  movel([0.295202, -1.405507, -2.534956, -0.771926, 1.570796, 1.865998],accel_mss,speed_ms,0,blend_radius_m)
  movel([0.293033, -1.404298, -2.535858, -0.772233, 1.570796, 1.863829],accel_mss,speed_ms,0,blend_radius_m)
  movel([0.292106, -1.403830, -2.536207, -0.772352, 1.570796, 1.862902],accel_mss,speed_ms,0,blend_radius_m)
  movel([0.292065, -1.403853, -2.536190, -0.772346, 1.570796, 1.862862],accel_mss,speed_ms,0,blend_radius_m)
  movel([0.291975, -1.403947, -2.536120, -0.772322, 1.570796, 1.862771],accel_mss,speed_ms,0,blend_radius_m)
  movel([0.291907, -1.404050, -2.536043, -0.772296, 1.570796, 1.862703],accel_mss,speed_ms,0,blend_radius_m)
  movel([0.288768, -1.410063, -2.531537, -0.770789, 1.570796, 1.859564],accel_mss,speed_ms,0,blend_radius_m)
  movel([0.288784, -1.410109, -2.531502, -0.770777, 1.570796, 1.859580],accel_mss,speed_ms,0,blend_radius_m)
  movel([0.288827, -1.410120, -2.531495, -0.770775, 1.570796, 1.859623],accel_mss,speed_ms,0,blend_radius_m)
  movel([0.296146, -1.408109, -2.533007, -0.771273, 1.570796, 1.866942],accel_mss,speed_ms,0,blend_radius_m)
  movel([0.296784, -1.407940, -2.533134, -0.771315, 1.570796, 1.867580],accel_mss,speed_ms,0,blend_radius_m)
  movel([0.297418, -1.407780, -2.533254, -0.771355, 1.570796, 1.868215],accel_mss,speed_ms,0,blend_radius_m)
  movel([0.297807, -1.407689, -2.533323, -0.771378, 1.570796, 1.868604],accel_mss,speed_ms,0,blend_radius_m)
  movel([0.298196, -1.407603, -2.533387, -0.771399, 1.570796, 1.868993],accel_mss,speed_ms,0,blend_radius_m)
  movel([0.298230, -1.407602, -2.533388, -0.771399, 1.570796, 1.869026],accel_mss,speed_ms,0,blend_radius_m)
  movel([0.298257, -1.407614, -2.533378, -0.771396, 1.570796, 1.869053],accel_mss,speed_ms,0,blend_radius_m)
  movel([0.298268, -1.407641, -2.533359, -0.771390, 1.570796, 1.869065],accel_mss,speed_ms,0,blend_radius_m)
  movel([0.298265, -1.407672, -2.533335, -0.771382, 1.570796, 1.869061],accel_mss,speed_ms,0,blend_radius_m)
  movel([0.298217, -1.407806, -2.533235, -0.771348, 1.570796, 1.869013],accel_mss,speed_ms,0,blend_radius_m)
  movel([0.298155, -1.407940, -2.533134, -0.771315, 1.570796, 1.868951],accel_mss,speed_ms,0,blend_radius_m)
  movel([0.298085, -1.408074, -2.533034, -0.771281, 1.570796, 1.868881],accel_mss,speed_ms,0,blend_radius_m)
  movel([0.296508, -1.410799, -2.530982, -0.770608, 1.570796, 1.867304],accel_mss,speed_ms,0,blend_radius_m)
  movel([0.294863, -1.413645, -2.528828, -0.769916, 1.570796, 1.865659],accel_mss,speed_ms,0,blend_radius_m)
  movel([0.294838, -1.413674, -2.528806, -0.769909, 1.570796, 1.865634],accel_mss,speed_ms,0,blend_radius_m)
  movel([0.294807, -1.413696, -2.528790, -0.769904, 1.570796, 1.865603],accel_mss,speed_ms,0,blend_radius_m)
  movel([0.294773, -1.413705, -2.528783, -0.769901, 1.570796, 1.865569],accel_mss,speed_ms,0,blend_radius_m)
  movel([0.292403, -1.414377, -2.528272, -0.769740, 1.570796, 1.863199],accel_mss,speed_ms,0,blend_radius_m)
  speed_ms = 0.003
  movel([0.292403, -1.402314, -2.522404, -0.787670, 1.570796, 1.863199],accel_mss,speed_ms,0,blend_radius_m)
  speed_ms = 0.01
  movel([0.292403, -1.379125, -2.510287, -0.822977, 1.570796, 1.863199],accel_mss,speed_ms,0,blend_radius_m)
  movel([0.317529, -1.353731, -2.528171, -0.830488, 1.570796, 1.888326],accel_mss,speed_ms,0,blend_radius_m)
  movel([0.317529, -1.377341, -2.540600, -0.794448, 1.570796, 1.888326],accel_mss,speed_ms,0,blend_radius_m)
  speed_ms = 0.003
  movel([0.317529, -1.386537, -2.545131, -0.780721, 1.570796, 1.888326],accel_mss,speed_ms,0,blend_radius_m)
  speed_ms = 0.007
  movel([0.317400, -1.386449, -2.545195, -0.780745, 1.570796, 1.888196],accel_mss,speed_ms,0,blend_radius_m)
  movel([0.317282, -1.386351, -2.545265, -0.780773, 1.570796, 1.888079],accel_mss,speed_ms,0,blend_radius_m)
  movel([0.317179, -1.386239, -2.545346, -0.780804, 1.570796, 1.887975],accel_mss,speed_ms,0,blend_radius_m)
  movel([0.317088, -1.386117, -2.545434, -0.780838, 1.570796, 1.887884],accel_mss,speed_ms,0,blend_radius_m)
  movel([0.317009, -1.385985, -2.545529, -0.780875, 1.570796, 1.887805],accel_mss,speed_ms,0,blend_radius_m)
  movel([0.316947, -1.385844, -2.545630, -0.780915, 1.570796, 1.887743],accel_mss,speed_ms,0,blend_radius_m)
  movel([0.316895, -1.385687, -2.545744, -0.780959, 1.570796, 1.887691],accel_mss,speed_ms,0,blend_radius_m)
  movel([0.316856, -1.385524, -2.545861, -0.781004, 1.570796, 1.887652],accel_mss,speed_ms,0,blend_radius_m)
  movel([0.316831, -1.385353, -2.545983, -0.781052, 1.570796, 1.887627],accel_mss,speed_ms,0,blend_radius_m)
  movel([0.316820, -1.385175, -2.546111, -0.781102, 1.570796, 1.887616],accel_mss,speed_ms,0,blend_radius_m)
  movel([0.316821, -1.384994, -2.546242, -0.781153, 1.570796, 1.887617],accel_mss,speed_ms,0,blend_radius_m)
  movel([0.316837, -1.384809, -2.546374, -0.781205, 1.570796, 1.887633],accel_mss,speed_ms,0,blend_radius_m)
  movel([0.316871, -1.384610, -2.546517, -0.781261, 1.570796, 1.887668],accel_mss,speed_ms,0,blend_radius_m)
  movel([0.316923, -1.384407, -2.546663, -0.781318, 1.570796, 1.887719],accel_mss,speed_ms,0,blend_radius_m)
  movel([0.316994, -1.384201, -2.546811, -0.781377, 1.570796, 1.887790],accel_mss,speed_ms,0,blend_radius_m)
  movel([0.317085, -1.383995, -2.546959, -0.781435, 1.570796, 1.887881],accel_mss,speed_ms,0,blend_radius_m)
  movel([0.317196, -1.383778, -2.547115, -0.781496, 1.570796, 1.887992],accel_mss,speed_ms,0,blend_radius_m)
  movel([0.317324, -1.383562, -2.547269, -0.781557, 1.570796, 1.888120],accel_mss,speed_ms,0,blend_radius_m)
  movel([0.317466, -1.383347, -2.547423, -0.781618, 1.570796, 1.888262],accel_mss,speed_ms,0,blend_radius_m)
  movel([0.317621, -1.383138, -2.547573, -0.781678, 1.570796, 1.888418],accel_mss,speed_ms,0,blend_radius_m)
  movel([0.317789, -1.382934, -2.547719, -0.781736, 1.570796, 1.888585],accel_mss,speed_ms,0,blend_radius_m)
  movel([0.317971, -1.382735, -2.547862, -0.781792, 1.570796, 1.888767],accel_mss,speed_ms,0,blend_radius_m)
  movel([0.318163, -1.382544, -2.547998, -0.781847, 1.570796, 1.888959],accel_mss,speed_ms,0,blend_radius_m)
  movel([0.318364, -1.382361, -2.548129, -0.781899, 1.570796, 1.889161],accel_mss,speed_ms,0,blend_radius_m)
  movel([0.318563, -1.382197, -2.548246, -0.781946, 1.570796, 1.889360],accel_mss,speed_ms,0,blend_radius_m)
  movel([0.318773, -1.382043, -2.548356, -0.781989, 1.570796, 1.889569],accel_mss,speed_ms,0,blend_radius_m)
  movel([0.318988, -1.381904, -2.548455, -0.782029, 1.570796, 1.889784],accel_mss,speed_ms,0,blend_radius_m)
  movel([0.319211, -1.381778, -2.548546, -0.782065, 1.570796, 1.890007],accel_mss,speed_ms,0,blend_radius_m)
  movel([0.319370, -1.381698, -2.548603, -0.782088, 1.570796, 1.890166],accel_mss,speed_ms,0,blend_radius_m)
  movel([0.319528, -1.381626, -2.548654, -0.782109, 1.570796, 1.890324],accel_mss,speed_ms,0,blend_radius_m)
  movel([0.319666, -1.381574, -2.548691, -0.782124, 1.570796, 1.890463],accel_mss,speed_ms,0,blend_radius_m)
  movel([0.319802, -1.381535, -2.548719, -0.782135, 1.570796, 1.890598],accel_mss,speed_ms,0,blend_radius_m)
  movel([0.319954, -1.381503, -2.548742, -0.782144, 1.570796, 1.890750],accel_mss,speed_ms,0,blend_radius_m)
  movel([0.320103, -1.381485, -2.548755, -0.782149, 1.570796, 1.890899],accel_mss,speed_ms,0,blend_radius_m)
  movel([0.320317, -1.381467, -2.548768, -0.782154, 1.570796, 1.891114],accel_mss,speed_ms,0,blend_radius_m)
  movel([0.320529, -1.381457, -2.548775, -0.782157, 1.570796, 1.891326],accel_mss,speed_ms,0,blend_radius_m)
  movel([0.320739, -1.381453, -2.548778, -0.782158, 1.570796, 1.891535],accel_mss,speed_ms,0,blend_radius_m)
  movel([0.320944, -1.381456, -2.548776, -0.782157, 1.570796, 1.891740],accel_mss,speed_ms,0,blend_radius_m)
  movel([0.321088, -1.381466, -2.548768, -0.782154, 1.570796, 1.891884],accel_mss,speed_ms,0,blend_radius_m)
  movel([0.321225, -1.381490, -2.548751, -0.782148, 1.570796, 1.892021],accel_mss,speed_ms,0,blend_radius_m)
  movel([0.321339, -1.381527, -2.548725, -0.782137, 1.570796, 1.892135],accel_mss,speed_ms,0,blend_radius_m)
  movel([0.321447, -1.381575, -2.548691, -0.782123, 1.570796, 1.892243],accel_mss,speed_ms,0,blend_radius_m)
  movel([0.321565, -1.381645, -2.548640, -0.782103, 1.570796, 1.892361],accel_mss,speed_ms,0,blend_radius_m)
  movel([0.321678, -1.381723, -2.548585, -0.782081, 1.570796, 1.892474],accel_mss,speed_ms,0,blend_radius_m)
  movel([0.321782, -1.381815, -2.548519, -0.782055, 1.570796, 1.892578],accel_mss,speed_ms,0,blend_radius_m)
  movel([0.321874, -1.381914, -2.548449, -0.782026, 1.570796, 1.892671],accel_mss,speed_ms,0,blend_radius_m)
  movel([0.321956, -1.382025, -2.548370, -0.781995, 1.570796, 1.892752],accel_mss,speed_ms,0,blend_radius_m)
  movel([0.322026, -1.382143, -2.548285, -0.781961, 1.570796, 1.892822],accel_mss,speed_ms,0,blend_radius_m)
  movel([0.322084, -1.382268, -2.548195, -0.781925, 1.570796, 1.892880],accel_mss,speed_ms,0,blend_radius_m)
  movel([0.322142, -1.382446, -2.548068, -0.781875, 1.570796, 1.892938],accel_mss,speed_ms,0,blend_radius_m)
  movel([0.322181, -1.382631, -2.547936, -0.781822, 1.570796, 1.892978],accel_mss,speed_ms,0,blend_radius_m)
  movel([0.322201, -1.382827, -2.547796, -0.781766, 1.570796, 1.892998],accel_mss,speed_ms,0,blend_radius_m)
  movel([0.322206, -1.383028, -2.547652, -0.781709, 1.570796, 1.893002],accel_mss,speed_ms,0,blend_radius_m)
  movel([0.322190, -1.383244, -2.547497, -0.781648, 1.570796, 1.892986],accel_mss,speed_ms,0,blend_radius_m)
  movel([0.322153, -1.383466, -2.547339, -0.781585, 1.570796, 1.892949],accel_mss,speed_ms,0,blend_radius_m)
  movel([0.322100, -1.383688, -2.547179, -0.781522, 1.570796, 1.892897],accel_mss,speed_ms,0,blend_radius_m)
  movel([0.322031, -1.383914, -2.547017, -0.781458, 1.570796, 1.892827],accel_mss,speed_ms,0,blend_radius_m)
  movel([0.321941, -1.384144, -2.546852, -0.781393, 1.570796, 1.892738],accel_mss,speed_ms,0,blend_radius_m)
  movel([0.321837, -1.384373, -2.546688, -0.781328, 1.570796, 1.892633],accel_mss,speed_ms,0,blend_radius_m)
  movel([0.321714, -1.384603, -2.546523, -0.781263, 1.570796, 1.892510],accel_mss,speed_ms,0,blend_radius_m)
  movel([0.321577, -1.384828, -2.546361, -0.781200, 1.570796, 1.892373],accel_mss,speed_ms,0,blend_radius_m)
  movel([0.321470, -1.384985, -2.546248, -0.781156, 1.570796, 1.892267],accel_mss,speed_ms,0,blend_radius_m)
  movel([0.321350, -1.385137, -2.546139, -0.781113, 1.570796, 1.892146],accel_mss,speed_ms,0,blend_radius_m)
  movel([0.321218, -1.385283, -2.546034, -0.781072, 1.570796, 1.892014],accel_mss,speed_ms,0,blend_radius_m)
  movel([0.321054, -1.385449, -2.545914, -0.781025, 1.570796, 1.891850],accel_mss,speed_ms,0,blend_radius_m)
  movel([0.320882, -1.385612, -2.545798, -0.780980, 1.570796, 1.891679],accel_mss,speed_ms,0,blend_radius_m)
  movel([0.320704, -1.385768, -2.545685, -0.780936, 1.570796, 1.891500],accel_mss,speed_ms,0,blend_radius_m)
  movel([0.320519, -1.385918, -2.545577, -0.780894, 1.570796, 1.891315],accel_mss,speed_ms,0,blend_radius_m)
  movel([0.320332, -1.386060, -2.545475, -0.780854, 1.570796, 1.891128],accel_mss,speed_ms,0,blend_radius_m)
  movel([0.320137, -1.386198, -2.545375, -0.780815, 1.570796, 1.890934],accel_mss,speed_ms,0,blend_radius_m)
  movel([0.319967, -1.386307, -2.545297, -0.780785, 1.570796, 1.890763],accel_mss,speed_ms,0,blend_radius_m)
  movel([0.319794, -1.386402, -2.545228, -0.780759, 1.570796, 1.890590],accel_mss,speed_ms,0,blend_radius_m)
  movel([0.319615, -1.386489, -2.545165, -0.780734, 1.570796, 1.890411],accel_mss,speed_ms,0,blend_radius_m)
  movel([0.319423, -1.386569, -2.545108, -0.780712, 1.570796, 1.890219],accel_mss,speed_ms,0,blend_radius_m)
  movel([0.319229, -1.386634, -2.545061, -0.780694, 1.570796, 1.890026],accel_mss,speed_ms,0,blend_radius_m)
  movel([0.319037, -1.386688, -2.545022, -0.780679, 1.570796, 1.889833],accel_mss,speed_ms,0,blend_radius_m)
  movel([0.318848, -1.386727, -2.544994, -0.780668, 1.570796, 1.889644],accel_mss,speed_ms,0,blend_radius_m)
  movel([0.318659, -1.386753, -2.544976, -0.780661, 1.570796, 1.889455],accel_mss,speed_ms,0,blend_radius_m)
  movel([0.318477, -1.386763, -2.544968, -0.780658, 1.570796, 1.889273],accel_mss,speed_ms,0,blend_radius_m)
  movel([0.318298, -1.386760, -2.544970, -0.780659, 1.570796, 1.889094],accel_mss,speed_ms,0,blend_radius_m)
  movel([0.318128, -1.386741, -2.544984, -0.780664, 1.570796, 1.888925],accel_mss,speed_ms,0,blend_radius_m)
  movel([0.317963, -1.386711, -2.545005, -0.780672, 1.570796, 1.888759],accel_mss,speed_ms,0,blend_radius_m)
  movel([0.317810, -1.386666, -2.545038, -0.780685, 1.570796, 1.888606],accel_mss,speed_ms,0,blend_radius_m)
  movel([0.317665, -1.386608, -2.545080, -0.780701, 1.570796, 1.888461],accel_mss,speed_ms,0,blend_radius_m)
  movel([0.317529, -1.386537, -2.545131, -0.780721, 1.570796, 1.888326],accel_mss,speed_ms,0,blend_radius_m)
  speed_ms = 0.003
  movel([0.317529, -1.389645, -2.546625, -0.776120, 1.570796, 1.888326],accel_mss,speed_ms,0,blend_radius_m)
  speed_ms = 0.007
  movel([0.317400, -1.389556, -2.546689, -0.776144, 1.570796, 1.888196],accel_mss,speed_ms,0,blend_radius_m)
  movel([0.317282, -1.389458, -2.546760, -0.776171, 1.570796, 1.888079],accel_mss,speed_ms,0,blend_radius_m)
  movel([0.317179, -1.389346, -2.546841, -0.776202, 1.570796, 1.887975],accel_mss,speed_ms,0,blend_radius_m)
  movel([0.317088, -1.389225, -2.546929, -0.776235, 1.570796, 1.887884],accel_mss,speed_ms,0,blend_radius_m)
  movel([0.317009, -1.389094, -2.547024, -0.776272, 1.570796, 1.887805],accel_mss,speed_ms,0,blend_radius_m)
  movel([0.316947, -1.388953, -2.547126, -0.776311, 1.570796, 1.887743],accel_mss,speed_ms,0,blend_radius_m)
  movel([0.316895, -1.388796, -2.547239, -0.776354, 1.570796, 1.887691],accel_mss,speed_ms,0,blend_radius_m)
  movel([0.316856, -1.388633, -2.547356, -0.776399, 1.570796, 1.887652],accel_mss,speed_ms,0,blend_radius_m)
  movel([0.316831, -1.388463, -2.547479, -0.776446, 1.570796, 1.887627],accel_mss,speed_ms,0,blend_radius_m)
  movel([0.316820, -1.388286, -2.547608, -0.776496, 1.570796, 1.887616],accel_mss,speed_ms,0,blend_radius_m)
  movel([0.316821, -1.388105, -2.547738, -0.776546, 1.570796, 1.887617],accel_mss,speed_ms,0,blend_radius_m)
  movel([0.316837, -1.387921, -2.547871, -0.776597, 1.570796, 1.887633],accel_mss,speed_ms,0,blend_radius_m)
  movel([0.316871, -1.387722, -2.548015, -0.776652, 1.570796, 1.887668],accel_mss,speed_ms,0,blend_radius_m)
  movel([0.316923, -1.387520, -2.548160, -0.776709, 1.570796, 1.887719],accel_mss,speed_ms,0,blend_radius_m)
  movel([0.316994, -1.387314, -2.548309, -0.776766, 1.570796, 1.887790],accel_mss,speed_ms,0,blend_radius_m)
  movel([0.317085, -1.387108, -2.548457, -0.776824, 1.570796, 1.887881],accel_mss,speed_ms,0,blend_radius_m)
  movel([0.317196, -1.386892, -2.548613, -0.776884, 1.570796, 1.887992],accel_mss,speed_ms,0,blend_radius_m)
  movel([0.317324, -1.386677, -2.548768, -0.776944, 1.570796, 1.888120],accel_mss,speed_ms,0,blend_radius_m)
  movel([0.317466, -1.386462, -2.548922, -0.777004, 1.570796, 1.888262],accel_mss,speed_ms,0,blend_radius_m)
  movel([0.317621, -1.386253, -2.549073, -0.777063, 1.570796, 1.888418],accel_mss,speed_ms,0,blend_radius_m)
  movel([0.317789, -1.386050, -2.549219, -0.777120, 1.570796, 1.888585],accel_mss,speed_ms,0,blend_radius_m)
  movel([0.317971, -1.385851, -2.549362, -0.777176, 1.570796, 1.888767],accel_mss,speed_ms,0,blend_radius_m)
  movel([0.318163, -1.385661, -2.549499, -0.777229, 1.570796, 1.888959],accel_mss,speed_ms,0,blend_radius_m)
  movel([0.318364, -1.385478, -2.549630, -0.777281, 1.570796, 1.889161],accel_mss,speed_ms,0,blend_radius_m)
  movel([0.318563, -1.385315, -2.549747, -0.777327, 1.570796, 1.889360],accel_mss,speed_ms,0,blend_radius_m)
  movel([0.318773, -1.385162, -2.549857, -0.777370, 1.570796, 1.889569],accel_mss,speed_ms,0,blend_radius_m)
  movel([0.318988, -1.385023, -2.549957, -0.777409, 1.570796, 1.889784],accel_mss,speed_ms,0,blend_radius_m)
  movel([0.319211, -1.384897, -2.550047, -0.777445, 1.570796, 1.890007],accel_mss,speed_ms,0,blend_radius_m)
  movel([0.319370, -1.384817, -2.550105, -0.777467, 1.570796, 1.890166],accel_mss,speed_ms,0,blend_radius_m)
  movel([0.319528, -1.384746, -2.550156, -0.777488, 1.570796, 1.890324],accel_mss,speed_ms,0,blend_radius_m)
  movel([0.319666, -1.384693, -2.550193, -0.777502, 1.570796, 1.890463],accel_mss,speed_ms,0,blend_radius_m)
  movel([0.319802, -1.384654, -2.550221, -0.777513, 1.570796, 1.890598],accel_mss,speed_ms,0,blend_radius_m)
  movel([0.319954, -1.384623, -2.550244, -0.777522, 1.570796, 1.890750],accel_mss,speed_ms,0,blend_radius_m)
  movel([0.320103, -1.384604, -2.550257, -0.777528, 1.570796, 1.890899],accel_mss,speed_ms,0,blend_radius_m)
  movel([0.320317, -1.384587, -2.550270, -0.777532, 1.570796, 1.891114],accel_mss,speed_ms,0,blend_radius_m)
  movel([0.320529, -1.384576, -2.550277, -0.777535, 1.570796, 1.891326],accel_mss,speed_ms,0,blend_radius_m)
  movel([0.320739, -1.384573, -2.550280, -0.777537, 1.570796, 1.891535],accel_mss,speed_ms,0,blend_radius_m)
  movel([0.320944, -1.384576, -2.550278, -0.777536, 1.570796, 1.891740],accel_mss,speed_ms,0,blend_radius_m)
  movel([0.321088, -1.384586, -2.550270, -0.777533, 1.570796, 1.891884],accel_mss,speed_ms,0,blend_radius_m)
  movel([0.321225, -1.384610, -2.550253, -0.777526, 1.570796, 1.892021],accel_mss,speed_ms,0,blend_radius_m)
  movel([0.321339, -1.384646, -2.550227, -0.777516, 1.570796, 1.892135],accel_mss,speed_ms,0,blend_radius_m)
  movel([0.321447, -1.384694, -2.550193, -0.777502, 1.570796, 1.892243],accel_mss,speed_ms,0,blend_radius_m)
  movel([0.321565, -1.384765, -2.550142, -0.777482, 1.570796, 1.892361],accel_mss,speed_ms,0,blend_radius_m)
  movel([0.321678, -1.384842, -2.550086, -0.777460, 1.570796, 1.892474],accel_mss,speed_ms,0,blend_radius_m)
  movel([0.321782, -1.384934, -2.550021, -0.777434, 1.570796, 1.892578],accel_mss,speed_ms,0,blend_radius_m)
  movel([0.321874, -1.385032, -2.549950, -0.777407, 1.570796, 1.892671],accel_mss,speed_ms,0,blend_radius_m)
  movel([0.321956, -1.385143, -2.549871, -0.777375, 1.570796, 1.892752],accel_mss,speed_ms,0,blend_radius_m)
  movel([0.322026, -1.385261, -2.549786, -0.777342, 1.570796, 1.892822],accel_mss,speed_ms,0,blend_radius_m)
  movel([0.322084, -1.385386, -2.549696, -0.777307, 1.570796, 1.892880],accel_mss,speed_ms,0,blend_radius_m)
  movel([0.322142, -1.385563, -2.549569, -0.777257, 1.570796, 1.892938],accel_mss,speed_ms,0,blend_radius_m)
  movel([0.322181, -1.385748, -2.549436, -0.777205, 1.570796, 1.892978],accel_mss,speed_ms,0,blend_radius_m)
  movel([0.322201, -1.385943, -2.549296, -0.777150, 1.570796, 1.892998],accel_mss,speed_ms,0,blend_radius_m)
  movel([0.322206, -1.386144, -2.549151, -0.777094, 1.570796, 1.893002],accel_mss,speed_ms,0,blend_radius_m)
  movel([0.322190, -1.386359, -2.548997, -0.777033, 1.570796, 1.892986],accel_mss,speed_ms,0,blend_radius_m)
  movel([0.322153, -1.386580, -2.548837, -0.776971, 1.570796, 1.892949],accel_mss,speed_ms,0,blend_radius_m)
  movel([0.322100, -1.386802, -2.548677, -0.776909, 1.570796, 1.892897],accel_mss,speed_ms,0,blend_radius_m)
  movel([0.322031, -1.387028, -2.548515, -0.776846, 1.570796, 1.892827],accel_mss,speed_ms,0,blend_radius_m)
  movel([0.321941, -1.387257, -2.548350, -0.776782, 1.570796, 1.892738],accel_mss,speed_ms,0,blend_radius_m)
  movel([0.321837, -1.387485, -2.548185, -0.776718, 1.570796, 1.892633],accel_mss,speed_ms,0,blend_radius_m)
  movel([0.321714, -1.387715, -2.548020, -0.776654, 1.570796, 1.892510],accel_mss,speed_ms,0,blend_radius_m)
  movel([0.321577, -1.387939, -2.547858, -0.776592, 1.570796, 1.892373],accel_mss,speed_ms,0,blend_radius_m)
  movel([0.321470, -1.388096, -2.547745, -0.776548, 1.570796, 1.892267],accel_mss,speed_ms,0,blend_radius_m)
  movel([0.321350, -1.388248, -2.547635, -0.776506, 1.570796, 1.892146],accel_mss,speed_ms,0,blend_radius_m)
  movel([0.321218, -1.388393, -2.547530, -0.776466, 1.570796, 1.892014],accel_mss,speed_ms,0,blend_radius_m)
  movel([0.321054, -1.388559, -2.547410, -0.776420, 1.570796, 1.891850],accel_mss,speed_ms,0,blend_radius_m)
  movel([0.320882, -1.388721, -2.547293, -0.776375, 1.570796, 1.891679],accel_mss,speed_ms,0,blend_radius_m)
  movel([0.320704, -1.388877, -2.547180, -0.776332, 1.570796, 1.891500],accel_mss,speed_ms,0,blend_radius_m)
  movel([0.320519, -1.389027, -2.547072, -0.776290, 1.570796, 1.891315],accel_mss,speed_ms,0,blend_radius_m)
  movel([0.320332, -1.389169, -2.546969, -0.776251, 1.570796, 1.891128],accel_mss,speed_ms,0,blend_radius_m)
  movel([0.320137, -1.389306, -2.546870, -0.776213, 1.570796, 1.890934],accel_mss,speed_ms,0,blend_radius_m)
  movel([0.319967, -1.389414, -2.546792, -0.776183, 1.570796, 1.890763],accel_mss,speed_ms,0,blend_radius_m)
  movel([0.319794, -1.389510, -2.546723, -0.776157, 1.570796, 1.890590],accel_mss,speed_ms,0,blend_radius_m)
  movel([0.319615, -1.389597, -2.546660, -0.776133, 1.570796, 1.890411],accel_mss,speed_ms,0,blend_radius_m)
  movel([0.319423, -1.389676, -2.546602, -0.776111, 1.570796, 1.890219],accel_mss,speed_ms,0,blend_radius_m)
  movel([0.319229, -1.389741, -2.546555, -0.776093, 1.570796, 1.890026],accel_mss,speed_ms,0,blend_radius_m)
  movel([0.319037, -1.389795, -2.546516, -0.776078, 1.570796, 1.889833],accel_mss,speed_ms,0,blend_radius_m)
  movel([0.318848, -1.389833, -2.546488, -0.776067, 1.570796, 1.889644],accel_mss,speed_ms,0,blend_radius_m)
  movel([0.318659, -1.389859, -2.546469, -0.776060, 1.570796, 1.889455],accel_mss,speed_ms,0,blend_radius_m)
  movel([0.318477, -1.389869, -2.546462, -0.776058, 1.570796, 1.889273],accel_mss,speed_ms,0,blend_radius_m)
  movel([0.318298, -1.389866, -2.546464, -0.776058, 1.570796, 1.889094],accel_mss,speed_ms,0,blend_radius_m)
  movel([0.318128, -1.389848, -2.546478, -0.776064, 1.570796, 1.888925],accel_mss,speed_ms,0,blend_radius_m)
  movel([0.317963, -1.389818, -2.546499, -0.776072, 1.570796, 1.888759],accel_mss,speed_ms,0,blend_radius_m)
  movel([0.317810, -1.389772, -2.546532, -0.776084, 1.570796, 1.888606],accel_mss,speed_ms,0,blend_radius_m)
  movel([0.317665, -1.389715, -2.546574, -0.776100, 1.570796, 1.888461],accel_mss,speed_ms,0,blend_radius_m)
  movel([0.317529, -1.389645, -2.546625, -0.776120, 1.570796, 1.888326],accel_mss,speed_ms,0,blend_radius_m)
  speed_ms = 0.003
  movel([0.317529, -1.377341, -2.540600, -0.794448, 1.570796, 1.888326],accel_mss,speed_ms,0,blend_radius_m)
  speed_ms = 0.01
  movel([0.317529, -1.353731, -2.528171, -0.830488, 1.570796, 1.888326],accel_mss,speed_ms,0,blend_radius_m)
  movel([0.299954, -1.366063, -2.519594, -0.826732, 1.570796, 1.870750],accel_mss,speed_ms,0,blend_radius_m)
  movel([0.299954, -1.389472, -2.531871, -0.791046, 1.570796, 1.870750],accel_mss,speed_ms,0,blend_radius_m)
  speed_ms = 0.003
  movel([0.299954, -1.398583, -2.536345, -0.777462, 1.570796, 1.870750],accel_mss,speed_ms,0,blend_radius_m)
  speed_ms = 0.007
  movel([0.299979, -1.398601, -2.536331, -0.777457, 1.570796, 1.870775],accel_mss,speed_ms,0,blend_radius_m)
  movel([0.299990, -1.398630, -2.536310, -0.777450, 1.570796, 1.870786],accel_mss,speed_ms,0,blend_radius_m)
  movel([0.299985, -1.398664, -2.536284, -0.777441, 1.570796, 1.870782],accel_mss,speed_ms,0,blend_radius_m)
  movel([0.299976, -1.398686, -2.536268, -0.777435, 1.570796, 1.870772],accel_mss,speed_ms,0,blend_radius_m)
  movel([0.299706, -1.399170, -2.535911, -0.777308, 1.570796, 1.870502],accel_mss,speed_ms,0,blend_radius_m)
  movel([0.299404, -1.399711, -2.535511, -0.777167, 1.570796, 1.870201],accel_mss,speed_ms,0,blend_radius_m)
  movel([0.299046, -1.400345, -2.535042, -0.777003, 1.570796, 1.869842],accel_mss,speed_ms,0,blend_radius_m)
  movel([0.298078, -1.402098, -2.533741, -0.776550, 1.570796, 1.868875],accel_mss,speed_ms,0,blend_radius_m)
  movel([0.298054, -1.402119, -2.533726, -0.776545, 1.570796, 1.868850],accel_mss,speed_ms,0,blend_radius_m)
  movel([0.298027, -1.402128, -2.533719, -0.776542, 1.570796, 1.868823],accel_mss,speed_ms,0,blend_radius_m)
  movel([0.298001, -1.402124, -2.533722, -0.776543, 1.570796, 1.868797],accel_mss,speed_ms,0,blend_radius_m)
  movel([0.297791, -1.402026, -2.533795, -0.776569, 1.570796, 1.868587],accel_mss,speed_ms,0,blend_radius_m)
  movel([0.297586, -1.401919, -2.533874, -0.776596, 1.570796, 1.868382],accel_mss,speed_ms,0,blend_radius_m)
  movel([0.297210, -1.401715, -2.534026, -0.776648, 1.570796, 1.868006],accel_mss,speed_ms,0,blend_radius_m)
  movel([0.296838, -1.401504, -2.534182, -0.776703, 1.570796, 1.867634],accel_mss,speed_ms,0,blend_radius_m)
  movel([0.294823, -1.400338, -2.535047, -0.777004, 1.570796, 1.865620],accel_mss,speed_ms,0,blend_radius_m)
  movel([0.291768, -1.398674, -2.536277, -0.777438, 1.570796, 1.862565],accel_mss,speed_ms,0,blend_radius_m)
  movel([0.291698, -1.398742, -2.536227, -0.777420, 1.570796, 1.862494],accel_mss,speed_ms,0,blend_radius_m)
  movel([0.291646, -1.398819, -2.536170, -0.777400, 1.570796, 1.862443],accel_mss,speed_ms,0,blend_radius_m)
  movel([0.286418, -1.408830, -2.528706, -0.774853, 1.570796, 1.857214],accel_mss,speed_ms,0,blend_radius_m)
  movel([0.286404, -1.408924, -2.528635, -0.774830, 1.570796, 1.857200],accel_mss,speed_ms,0,blend_radius_m)
  movel([0.286418, -1.408956, -2.528611, -0.774822, 1.570796, 1.857214],accel_mss,speed_ms,0,blend_radius_m)
  movel([0.286461, -1.408960, -2.528608, -0.774821, 1.570796, 1.857257],accel_mss,speed_ms,0,blend_radius_m)
  movel([0.289039, -1.408279, -2.529120, -0.774990, 1.570796, 1.859835],accel_mss,speed_ms,0,blend_radius_m)
  movel([0.292788, -1.407230, -2.529908, -0.775251, 1.570796, 1.863584],accel_mss,speed_ms,0,blend_radius_m)
  movel([0.294307, -1.406809, -2.530224, -0.775356, 1.570796, 1.865103],accel_mss,speed_ms,0,blend_radius_m)
  movel([0.295651, -1.406440, -2.530501, -0.775448, 1.570796, 1.866448],accel_mss,speed_ms,0,blend_radius_m)
  movel([0.295756, -1.406418, -2.530517, -0.775454, 1.570796, 1.866552],accel_mss,speed_ms,0,blend_radius_m)
  movel([0.295779, -1.406422, -2.530514, -0.775453, 1.570796, 1.866575],accel_mss,speed_ms,0,blend_radius_m)
  movel([0.295789, -1.406438, -2.530502, -0.775449, 1.570796, 1.866585],accel_mss,speed_ms,0,blend_radius_m)
  movel([0.295786, -1.406461, -2.530485, -0.775443, 1.570796, 1.866582],accel_mss,speed_ms,0,blend_radius_m)
  movel([0.295610, -1.406827, -2.530211, -0.775351, 1.570796, 1.866406],accel_mss,speed_ms,0,blend_radius_m)
  movel([0.295483, -1.407076, -2.530024, -0.775289, 1.570796, 1.866279],accel_mss,speed_ms,0,blend_radius_m)
  movel([0.295348, -1.407323, -2.529838, -0.775227, 1.570796, 1.866144],accel_mss,speed_ms,0,blend_radius_m)
  movel([0.294960, -1.408010, -2.529323, -0.775057, 1.570796, 1.865757],accel_mss,speed_ms,0,blend_radius_m)
  movel([0.294039, -1.409616, -2.528114, -0.774660, 1.570796, 1.864835],accel_mss,speed_ms,0,blend_radius_m)
  movel([0.286883, -1.411688, -2.526548, -0.774153, 1.570796, 1.857680],accel_mss,speed_ms,0,blend_radius_m)
  movel([0.279741, -1.413793, -2.524951, -0.773645, 1.570796, 1.850537],accel_mss,speed_ms,0,blend_radius_m)
  movel([0.278382, -1.412114, -2.526226, -0.774050, 1.570796, 1.849178],accel_mss,speed_ms,0,blend_radius_m)
  movel([0.277016, -1.410434, -2.527496, -0.774459, 1.570796, 1.847813],accel_mss,speed_ms,0,blend_radius_m)
  movel([0.280791, -1.403859, -2.532430, -0.776100, 1.570796, 1.851587],accel_mss,speed_ms,0,blend_radius_m)
  movel([0.282261, -1.401314, -2.534323, -0.776752, 1.570796, 1.853058],accel_mss,speed_ms,0,blend_radius_m)
  movel([0.283526, -1.399146, -2.535928, -0.777314, 1.570796, 1.854322],accel_mss,speed_ms,0,blend_radius_m)
  movel([0.284665, -1.397209, -2.537357, -0.777823, 1.570796, 1.855461],accel_mss,speed_ms,0,blend_radius_m)
  movel([0.284701, -1.397159, -2.537394, -0.777836, 1.570796, 1.855497],accel_mss,speed_ms,0,blend_radius_m)
  movel([0.284746, -1.397114, -2.537427, -0.777848, 1.570796, 1.855542],accel_mss,speed_ms,0,blend_radius_m)
  movel([0.284807, -1.397067, -2.537461, -0.777860, 1.570796, 1.855604],accel_mss,speed_ms,0,blend_radius_m)
  movel([0.284875, -1.397031, -2.537488, -0.777870, 1.570796, 1.855671],accel_mss,speed_ms,0,blend_radius_m)
  movel([0.284943, -1.397005, -2.537507, -0.777877, 1.570796, 1.855740],accel_mss,speed_ms,0,blend_radius_m)
  movel([0.287618, -1.396223, -2.538082, -0.778084, 1.570796, 1.858414],accel_mss,speed_ms,0,blend_radius_m)
  movel([0.290146, -1.395495, -2.538617, -0.778278, 1.570796, 1.860943],accel_mss,speed_ms,0,blend_radius_m)
  movel([0.290337, -1.395446, -2.538653, -0.778291, 1.570796, 1.861133],accel_mss,speed_ms,0,blend_radius_m)
  movel([0.290526, -1.395407, -2.538681, -0.778301, 1.570796, 1.861322],accel_mss,speed_ms,0,blend_radius_m)
  movel([0.290711, -1.395380, -2.538701, -0.778308, 1.570796, 1.861508],accel_mss,speed_ms,0,blend_radius_m)
  movel([0.290805, -1.395375, -2.538705, -0.778309, 1.570796, 1.861601],accel_mss,speed_ms,0,blend_radius_m)
  movel([0.290892, -1.395381, -2.538700, -0.778308, 1.570796, 1.861689],accel_mss,speed_ms,0,blend_radius_m)
  movel([0.290971, -1.395402, -2.538685, -0.778302, 1.570796, 1.861767],accel_mss,speed_ms,0,blend_radius_m)
  movel([0.295448, -1.396969, -2.537534, -0.777886, 1.570796, 1.866244],accel_mss,speed_ms,0,blend_radius_m)
  movel([0.299954, -1.398583, -2.536345, -0.777462, 1.570796, 1.870750],accel_mss,speed_ms,0,blend_radius_m)
  speed_ms = 0.003
  movel([0.299954, -1.401660, -2.537819, -0.772910, 1.570796, 1.870750],accel_mss,speed_ms,0,blend_radius_m)
  speed_ms = 0.007
  movel([0.299979, -1.401679, -2.537806, -0.772905, 1.570796, 1.870775],accel_mss,speed_ms,0,blend_radius_m)
  movel([0.299990, -1.401707, -2.537785, -0.772898, 1.570796, 1.870786],accel_mss,speed_ms,0,blend_radius_m)
  movel([0.299985, -1.401741, -2.537759, -0.772889, 1.570796, 1.870782],accel_mss,speed_ms,0,blend_radius_m)
  movel([0.299976, -1.401763, -2.537743, -0.772883, 1.570796, 1.870772],accel_mss,speed_ms,0,blend_radius_m)
  movel([0.299706, -1.402245, -2.537385, -0.772759, 1.570796, 1.870502],accel_mss,speed_ms,0,blend_radius_m)
  movel([0.299404, -1.402785, -2.536984, -0.772620, 1.570796, 1.870201],accel_mss,speed_ms,0,blend_radius_m)
  movel([0.299046, -1.403418, -2.536514, -0.772458, 1.570796, 1.869842],accel_mss,speed_ms,0,blend_radius_m)
  movel([0.298078, -1.405166, -2.535211, -0.772012, 1.570796, 1.868875],accel_mss,speed_ms,0,blend_radius_m)
  movel([0.298054, -1.405187, -2.535195, -0.772007, 1.570796, 1.868850],accel_mss,speed_ms,0,blend_radius_m)
  movel([0.298027, -1.405196, -2.535188, -0.772005, 1.570796, 1.868823],accel_mss,speed_ms,0,blend_radius_m)
  movel([0.298001, -1.405192, -2.535191, -0.772006, 1.570796, 1.868797],accel_mss,speed_ms,0,blend_radius_m)
  movel([0.297791, -1.405094, -2.535264, -0.772030, 1.570796, 1.868587],accel_mss,speed_ms,0,blend_radius_m)
  movel([0.297586, -1.404988, -2.535344, -0.772057, 1.570796, 1.868382],accel_mss,speed_ms,0,blend_radius_m)
  movel([0.297210, -1.404784, -2.535496, -0.772109, 1.570796, 1.868006],accel_mss,speed_ms,0,blend_radius_m)
  movel([0.296838, -1.404574, -2.535652, -0.772163, 1.570796, 1.867634],accel_mss,speed_ms,0,blend_radius_m)
  movel([0.294823, -1.403410, -2.536519, -0.772459, 1.570796, 1.865620],accel_mss,speed_ms,0,blend_radius_m)
  movel([0.291768, -1.401751, -2.537752, -0.772886, 1.570796, 1.862565],accel_mss,speed_ms,0,blend_radius_m)
  movel([0.291698, -1.401819, -2.537701, -0.772869, 1.570796, 1.862494],accel_mss,speed_ms,0,blend_radius_m)
  movel([0.291646, -1.401895, -2.537645, -0.772849, 1.570796, 1.862443],accel_mss,speed_ms,0,blend_radius_m)
  movel([0.286418, -1.411881, -2.530165, -0.770343, 1.570796, 1.857214],accel_mss,speed_ms,0,blend_radius_m)
  movel([0.286404, -1.411976, -2.530093, -0.770320, 1.570796, 1.857200],accel_mss,speed_ms,0,blend_radius_m)
  movel([0.286418, -1.412007, -2.530069, -0.770313, 1.570796, 1.857214],accel_mss,speed_ms,0,blend_radius_m)
  movel([0.286461, -1.412011, -2.530066, -0.770312, 1.570796, 1.857257],accel_mss,speed_ms,0,blend_radius_m)
  movel([0.289039, -1.411332, -2.530580, -0.770477, 1.570796, 1.859835],accel_mss,speed_ms,0,blend_radius_m)
  movel([0.292788, -1.410286, -2.531370, -0.770734, 1.570796, 1.863584],accel_mss,speed_ms,0,blend_radius_m)
  movel([0.294307, -1.409865, -2.531686, -0.770837, 1.570796, 1.865103],accel_mss,speed_ms,0,blend_radius_m)
  movel([0.295651, -1.409498, -2.531963, -0.770928, 1.570796, 1.866448],accel_mss,speed_ms,0,blend_radius_m)
  movel([0.295756, -1.409476, -2.531980, -0.770934, 1.570796, 1.866552],accel_mss,speed_ms,0,blend_radius_m)
  movel([0.295779, -1.409480, -2.531977, -0.770933, 1.570796, 1.866575],accel_mss,speed_ms,0,blend_radius_m)
  movel([0.295789, -1.409495, -2.531965, -0.770929, 1.570796, 1.866585],accel_mss,speed_ms,0,blend_radius_m)
  movel([0.295786, -1.409519, -2.531947, -0.770923, 1.570796, 1.866582],accel_mss,speed_ms,0,blend_radius_m)
  movel([0.295610, -1.409884, -2.531673, -0.770833, 1.570796, 1.866406],accel_mss,speed_ms,0,blend_radius_m)
  movel([0.295483, -1.410132, -2.531485, -0.770772, 1.570796, 1.866279],accel_mss,speed_ms,0,blend_radius_m)
  movel([0.295348, -1.410379, -2.531299, -0.770711, 1.570796, 1.866144],accel_mss,speed_ms,0,blend_radius_m)
  movel([0.294960, -1.411063, -2.530783, -0.770543, 1.570796, 1.865757],accel_mss,speed_ms,0,blend_radius_m)
  movel([0.294039, -1.412665, -2.529571, -0.770153, 1.570796, 1.864835],accel_mss,speed_ms,0,blend_radius_m)
  movel([0.286883, -1.414733, -2.528002, -0.769654, 1.570796, 1.857680],accel_mss,speed_ms,0,blend_radius_m)
  movel([0.279741, -1.416832, -2.526402, -0.769155, 1.570796, 1.850537],accel_mss,speed_ms,0,blend_radius_m)
  movel([0.278382, -1.415157, -2.527679, -0.769553, 1.570796, 1.849178],accel_mss,speed_ms,0,blend_radius_m)
  movel([0.277016, -1.413481, -2.528953, -0.769955, 1.570796, 1.847813],accel_mss,speed_ms,0,blend_radius_m)
  movel([0.280791, -1.406923, -2.533897, -0.771569, 1.570796, 1.851587],accel_mss,speed_ms,0,blend_radius_m)
  movel([0.282261, -1.404384, -2.535794, -0.772211, 1.570796, 1.853058],accel_mss,speed_ms,0,blend_radius_m)
  movel([0.283526, -1.402222, -2.537402, -0.772765, 1.570796, 1.854322],accel_mss,speed_ms,0,blend_radius_m)
  movel([0.284665, -1.400289, -2.538834, -0.773265, 1.570796, 1.855461],accel_mss,speed_ms,0,blend_radius_m)
  movel([0.284701, -1.400239, -2.538871, -0.773278, 1.570796, 1.855497],accel_mss,speed_ms,0,blend_radius_m)
  movel([0.284746, -1.400195, -2.538904, -0.773290, 1.570796, 1.855542],accel_mss,speed_ms,0,blend_radius_m)
  movel([0.284807, -1.400148, -2.538938, -0.773302, 1.570796, 1.855604],accel_mss,speed_ms,0,blend_radius_m)
  movel([0.284875, -1.400112, -2.538965, -0.773312, 1.570796, 1.855671],accel_mss,speed_ms,0,blend_radius_m)
  movel([0.284943, -1.400086, -2.538985, -0.773318, 1.570796, 1.855740],accel_mss,speed_ms,0,blend_radius_m)
  movel([0.287618, -1.399306, -2.539561, -0.773522, 1.570796, 1.858414],accel_mss,speed_ms,0,blend_radius_m)
  movel([0.290146, -1.398580, -2.540097, -0.773713, 1.570796, 1.860943],accel_mss,speed_ms,0,blend_radius_m)
  movel([0.290337, -1.398531, -2.540133, -0.773726, 1.570796, 1.861133],accel_mss,speed_ms,0,blend_radius_m)
  movel([0.290526, -1.398493, -2.540161, -0.773736, 1.570796, 1.861322],accel_mss,speed_ms,0,blend_radius_m)
  movel([0.290711, -1.398465, -2.540181, -0.773743, 1.570796, 1.861508],accel_mss,speed_ms,0,blend_radius_m)
  movel([0.290805, -1.398460, -2.540185, -0.773744, 1.570796, 1.861601],accel_mss,speed_ms,0,blend_radius_m)
  movel([0.290892, -1.398466, -2.540180, -0.773743, 1.570796, 1.861689],accel_mss,speed_ms,0,blend_radius_m)
  movel([0.290971, -1.398487, -2.540164, -0.773737, 1.570796, 1.861767],accel_mss,speed_ms,0,blend_radius_m)
  movel([0.295448, -1.400050, -2.539011, -0.773328, 1.570796, 1.866244],accel_mss,speed_ms,0,blend_radius_m)
  movel([0.299954, -1.401660, -2.537819, -0.772910, 1.570796, 1.870750],accel_mss,speed_ms,0,blend_radius_m)
  speed_ms = 0.003
  movel([0.299954, -1.389472, -2.531871, -0.791046, 1.570796, 1.870750],accel_mss,speed_ms,0,blend_radius_m)
  speed_ms = 0.01
  movel([0.299954, -1.366063, -2.519594, -0.826732, 1.570796, 1.870750],accel_mss,speed_ms,0,blend_radius_m)
  movel([0.309412, -1.329808, -2.544234, -0.838348, 1.570796, 1.880209],accel_mss,speed_ms,0,blend_radius_m)
  movel([0.309412, -1.353793, -2.556962, -0.801634, 1.570796, 1.880209],accel_mss,speed_ms,0,blend_radius_m)
  speed_ms = 0.003
  movel([0.309412, -1.363150, -2.561605, -0.787634, 1.570796, 1.880209],accel_mss,speed_ms,0,blend_radius_m)
  speed_ms = 0.007
  movel([0.297723, -1.363243, -2.561541, -0.787605, 1.570796, 1.868520],accel_mss,speed_ms,0,blend_radius_m)
  movel([0.285995, -1.363475, -2.561381, -0.787532, 1.570796, 1.856791],accel_mss,speed_ms,0,blend_radius_m)
  movel([0.285952, -1.363472, -2.561384, -0.787534, 1.570796, 1.856748],accel_mss,speed_ms,0,blend_radius_m)
  movel([0.285916, -1.363458, -2.561393, -0.787538, 1.570796, 1.856713],accel_mss,speed_ms,0,blend_radius_m)
  movel([0.285886, -1.363438, -2.561407, -0.787544, 1.570796, 1.856682],accel_mss,speed_ms,0,blend_radius_m)
  movel([0.285881, -1.363423, -2.561417, -0.787549, 1.570796, 1.856677],accel_mss,speed_ms,0,blend_radius_m)
  movel([0.285883, -1.363403, -2.561431, -0.787555, 1.570796, 1.856679],accel_mss,speed_ms,0,blend_radius_m)
  movel([0.286224, -1.362510, -2.562045, -0.787834, 1.570796, 1.857020],accel_mss,speed_ms,0,blend_radius_m)
  movel([0.286612, -1.361507, -2.562734, -0.788148, 1.570796, 1.857408],accel_mss,speed_ms,0,blend_radius_m)
  movel([0.287081, -1.360318, -2.563548, -0.788523, 1.570796, 1.857877],accel_mss,speed_ms,0,blend_radius_m)
  movel([0.288314, -1.357214, -2.565665, -0.789509, 1.570796, 1.859110],accel_mss,speed_ms,0,blend_radius_m)
  movel([0.288787, -1.357208, -2.565669, -0.789511, 1.570796, 1.859583],accel_mss,speed_ms,0,blend_radius_m)
  movel([0.292493, -1.357128, -2.565724, -0.789537, 1.570796, 1.863289],accel_mss,speed_ms,0,blend_radius_m)
  movel([0.300718, -1.356988, -2.565819, -0.789582, 1.570796, 1.871514],accel_mss,speed_ms,0,blend_radius_m)
  movel([0.312121, -1.356904, -2.565876, -0.789609, 1.570796, 1.882917],accel_mss,speed_ms,0,blend_radius_m)
  movel([0.312020, -1.357204, -2.565672, -0.789513, 1.570796, 1.882816],accel_mss,speed_ms,0,blend_radius_m)
  movel([0.311964, -1.357358, -2.565568, -0.789464, 1.570796, 1.882760],accel_mss,speed_ms,0,blend_radius_m)
  movel([0.311875, -1.357574, -2.565420, -0.789394, 1.570796, 1.882671],accel_mss,speed_ms,0,blend_radius_m)
  movel([0.311772, -1.357812, -2.565258, -0.789318, 1.570796, 1.882568],accel_mss,speed_ms,0,blend_radius_m)
  movel([0.311669, -1.358037, -2.565105, -0.789247, 1.570796, 1.882465],accel_mss,speed_ms,0,blend_radius_m)
  movel([0.311422, -1.358566, -2.564745, -0.789078, 1.570796, 1.882218],accel_mss,speed_ms,0,blend_radius_m)
  movel([0.309918, -1.358722, -2.564638, -0.789028, 1.570796, 1.880714],accel_mss,speed_ms,0,blend_radius_m)
  movel([0.308373, -1.358921, -2.564503, -0.788965, 1.570796, 1.879169],accel_mss,speed_ms,0,blend_radius_m)
  movel([0.308340, -1.358969, -2.564470, -0.788950, 1.570796, 1.879137],accel_mss,speed_ms,0,blend_radius_m)
  movel([0.307920, -1.361123, -2.562997, -0.788269, 1.570796, 1.878717],accel_mss,speed_ms,0,blend_radius_m)
  movel([0.310504, -1.360769, -2.563240, -0.788380, 1.570796, 1.881300],accel_mss,speed_ms,0,blend_radius_m)
  movel([0.310037, -1.361915, -2.562454, -0.788020, 1.570796, 1.880834],accel_mss,speed_ms,0,blend_radius_m)
  movel([0.309853, -1.362357, -2.562150, -0.787882, 1.570796, 1.880649],accel_mss,speed_ms,0,blend_radius_m)
  movel([0.309691, -1.362737, -2.561889, -0.787763, 1.570796, 1.880487],accel_mss,speed_ms,0,blend_radius_m)
  movel([0.309545, -1.363064, -2.561664, -0.787661, 1.570796, 1.880341],accel_mss,speed_ms,0,blend_radius_m)
  movel([0.309530, -1.363087, -2.561648, -0.787653, 1.570796, 1.880326],accel_mss,speed_ms,0,blend_radius_m)
  movel([0.309511, -1.363109, -2.561633, -0.787647, 1.570796, 1.880308],accel_mss,speed_ms,0,blend_radius_m)
  movel([0.309479, -1.363130, -2.561619, -0.787640, 1.570796, 1.880275],accel_mss,speed_ms,0,blend_radius_m)
  movel([0.309446, -1.363144, -2.561609, -0.787636, 1.570796, 1.880243],accel_mss,speed_ms,0,blend_radius_m)
  movel([0.309412, -1.363150, -2.561605, -0.787634, 1.570796, 1.880209],accel_mss,speed_ms,0,blend_radius_m)
  speed_ms = 0.003
  movel([0.309412, -1.366314, -2.563137, -0.782939, 1.570796, 1.880209],accel_mss,speed_ms,0,blend_radius_m)
  speed_ms = 0.007
  movel([0.297723, -1.366407, -2.563072, -0.782910, 1.570796, 1.868520],accel_mss,speed_ms,0,blend_radius_m)
  movel([0.285995, -1.366638, -2.562912, -0.782839, 1.570796, 1.856791],accel_mss,speed_ms,0,blend_radius_m)
  movel([0.285952, -1.366634, -2.562915, -0.782840, 1.570796, 1.856748],accel_mss,speed_ms,0,blend_radius_m)
  movel([0.285916, -1.366621, -2.562924, -0.782844, 1.570796, 1.856713],accel_mss,speed_ms,0,blend_radius_m)
  movel([0.285886, -1.366601, -2.562938, -0.782850, 1.570796, 1.856682],accel_mss,speed_ms,0,blend_radius_m)
  movel([0.285881, -1.366586, -2.562948, -0.782855, 1.570796, 1.856677],accel_mss,speed_ms,0,blend_radius_m)
  movel([0.285883, -1.366566, -2.562962, -0.782861, 1.570796, 1.856679],accel_mss,speed_ms,0,blend_radius_m)
  movel([0.286224, -1.365675, -2.563578, -0.783136, 1.570796, 1.857020],accel_mss,speed_ms,0,blend_radius_m)
  movel([0.286612, -1.364674, -2.564268, -0.783447, 1.570796, 1.857408],accel_mss,speed_ms,0,blend_radius_m)
  movel([0.287081, -1.363488, -2.565085, -0.783817, 1.570796, 1.857877],accel_mss,speed_ms,0,blend_radius_m)
  movel([0.288314, -1.360392, -2.567206, -0.784791, 1.570796, 1.859110],accel_mss,speed_ms,0,blend_radius_m)
  movel([0.288787, -1.360386, -2.567210, -0.784793, 1.570796, 1.859583],accel_mss,speed_ms,0,blend_radius_m)
  movel([0.292493, -1.360306, -2.567265, -0.784818, 1.570796, 1.863289],accel_mss,speed_ms,0,blend_radius_m)
  movel([0.300718, -1.360166, -2.567360, -0.784863, 1.570796, 1.871514],accel_mss,speed_ms,0,blend_radius_m)
  movel([0.312121, -1.360082, -2.567418, -0.784889, 1.570796, 1.882917],accel_mss,speed_ms,0,blend_radius_m)
  movel([0.312020, -1.360382, -2.567213, -0.784794, 1.570796, 1.882816],accel_mss,speed_ms,0,blend_radius_m)
  movel([0.311964, -1.360535, -2.567109, -0.784746, 1.570796, 1.882760],accel_mss,speed_ms,0,blend_radius_m)
  movel([0.311875, -1.360751, -2.566961, -0.784677, 1.570796, 1.882671],accel_mss,speed_ms,0,blend_radius_m)
  movel([0.311772, -1.360988, -2.566798, -0.784602, 1.570796, 1.882568],accel_mss,speed_ms,0,blend_radius_m)
  movel([0.311669, -1.361212, -2.566645, -0.784532, 1.570796, 1.882465],accel_mss,speed_ms,0,blend_radius_m)
  movel([0.311422, -1.361740, -2.566284, -0.784365, 1.570796, 1.882218],accel_mss,speed_ms,0,blend_radius_m)
  movel([0.309918, -1.361896, -2.566177, -0.784316, 1.570796, 1.880714],accel_mss,speed_ms,0,blend_radius_m)
  movel([0.308373, -1.362094, -2.566041, -0.784254, 1.570796, 1.879169],accel_mss,speed_ms,0,blend_radius_m)
  movel([0.308340, -1.362142, -2.566008, -0.784239, 1.570796, 1.879137],accel_mss,speed_ms,0,blend_radius_m)
  movel([0.307920, -1.364291, -2.564532, -0.783566, 1.570796, 1.878717],accel_mss,speed_ms,0,blend_radius_m)
  movel([0.310504, -1.363938, -2.564775, -0.783676, 1.570796, 1.881300],accel_mss,speed_ms,0,blend_radius_m)
  movel([0.310037, -1.365081, -2.563987, -0.783320, 1.570796, 1.880834],accel_mss,speed_ms,0,blend_radius_m)
  movel([0.309853, -1.365522, -2.563683, -0.783183, 1.570796, 1.880649],accel_mss,speed_ms,0,blend_radius_m)
  movel([0.309691, -1.365901, -2.563421, -0.783066, 1.570796, 1.880487],accel_mss,speed_ms,0,blend_radius_m)
  movel([0.309545, -1.366228, -2.563196, -0.782965, 1.570796, 1.880341],accel_mss,speed_ms,0,blend_radius_m)
  movel([0.309530, -1.366251, -2.563180, -0.782958, 1.570796, 1.880326],accel_mss,speed_ms,0,blend_radius_m)
  movel([0.309511, -1.366273, -2.563165, -0.782951, 1.570796, 1.880308],accel_mss,speed_ms,0,blend_radius_m)
  movel([0.309479, -1.366294, -2.563150, -0.782945, 1.570796, 1.880275],accel_mss,speed_ms,0,blend_radius_m)
  movel([0.309446, -1.366308, -2.563140, -0.782941, 1.570796, 1.880243],accel_mss,speed_ms,0,blend_radius_m)
  movel([0.309412, -1.366314, -2.563137, -0.782939, 1.570796, 1.880209],accel_mss,speed_ms,0,blend_radius_m)
  speed_ms = 0.003
  movel([0.309412, -1.353793, -2.556962, -0.801634, 1.570796, 1.880209],accel_mss,speed_ms,0,blend_radius_m)
  speed_ms = 0.01
  movel([0.309412, -1.329808, -2.544234, -0.838348, 1.570796, 1.880209],accel_mss,speed_ms,0,blend_radius_m)
  movel([0.310290, -1.321918, -2.549368, -0.841103, 1.570796, 1.881086],accel_mss,speed_ms,0,blend_radius_m)
  movel([0.310290, -1.346022, -2.562195, -0.804172, 1.570796, 1.881086],accel_mss,speed_ms,0,blend_radius_m)
  speed_ms = 0.003
  movel([0.310290, -1.355431, -2.566876, -0.790083, 1.570796, 1.881086],accel_mss,speed_ms,0,blend_radius_m)
  speed_ms = 0.007
  movel([0.310214, -1.355447, -2.566864, -0.790077, 1.570796, 1.881011],accel_mss,speed_ms,0,blend_radius_m)
  movel([0.310141, -1.355452, -2.566861, -0.790076, 1.570796, 1.880937],accel_mss,speed_ms,0,blend_radius_m)
  movel([0.309901, -1.355452, -2.566861, -0.790076, 1.570796, 1.880697],accel_mss,speed_ms,0,blend_radius_m)
  movel([0.308940, -1.355441, -2.566869, -0.790079, 1.570796, 1.879736],accel_mss,speed_ms,0,blend_radius_m)
  movel([0.298968, -1.355552, -2.566794, -0.790044, 1.570796, 1.869764],accel_mss,speed_ms,0,blend_radius_m)
  movel([0.288662, -1.355768, -2.566647, -0.789974, 1.570796, 1.859458],accel_mss,speed_ms,0,blend_radius_m)
  movel([0.288310, -1.355795, -2.566629, -0.789965, 1.570796, 1.859107],accel_mss,speed_ms,0,blend_radius_m)
  movel([0.288264, -1.355794, -2.566629, -0.789966, 1.570796, 1.859060],accel_mss,speed_ms,0,blend_radius_m)
  movel([0.288229, -1.355778, -2.566640, -0.789971, 1.570796, 1.859025],accel_mss,speed_ms,0,blend_radius_m)
  movel([0.288203, -1.355748, -2.566661, -0.789980, 1.570796, 1.859000],accel_mss,speed_ms,0,blend_radius_m)
  movel([0.288192, -1.355709, -2.566687, -0.789993, 1.570796, 1.858988],accel_mss,speed_ms,0,blend_radius_m)
  movel([0.288195, -1.355640, -2.566734, -0.790015, 1.570796, 1.858991],accel_mss,speed_ms,0,blend_radius_m)
  movel([0.288208, -1.355570, -2.566782, -0.790038, 1.570796, 1.859004],accel_mss,speed_ms,0,blend_radius_m)
  movel([0.288279, -1.355325, -2.566947, -0.790117, 1.570796, 1.859075],accel_mss,speed_ms,0,blend_radius_m)
  movel([0.288342, -1.355139, -2.567073, -0.790177, 1.570796, 1.859138],accel_mss,speed_ms,0,blend_radius_m)
  movel([0.288415, -1.354950, -2.567201, -0.790238, 1.570796, 1.859211],accel_mss,speed_ms,0,blend_radius_m)
  movel([0.289451, -1.352376, -2.568938, -0.791074, 1.570796, 1.860248],accel_mss,speed_ms,0,blend_radius_m)
  movel([0.290662, -1.349390, -2.570943, -0.792056, 1.570796, 1.861458],accel_mss,speed_ms,0,blend_radius_m)
  movel([0.292076, -1.345926, -2.573253, -0.793210, 1.570796, 1.862872],accel_mss,speed_ms,0,blend_radius_m)
  movel([0.295785, -1.336892, -2.579201, -0.796296, 1.570796, 1.866581],accel_mss,speed_ms,0,blend_radius_m)
  movel([0.296446, -1.336847, -2.579230, -0.796312, 1.570796, 1.867242],accel_mss,speed_ms,0,blend_radius_m)
  movel([0.296887, -1.336823, -2.579246, -0.796320, 1.570796, 1.867683],accel_mss,speed_ms,0,blend_radius_m)
  movel([0.297322, -1.336815, -2.579251, -0.796323, 1.570796, 1.868119],accel_mss,speed_ms,0,blend_radius_m)
  movel([0.297751, -1.336820, -2.579248, -0.796321, 1.570796, 1.868548],accel_mss,speed_ms,0,blend_radius_m)
  movel([0.298232, -1.336842, -2.579234, -0.796314, 1.570796, 1.869029],accel_mss,speed_ms,0,blend_radius_m)
  movel([0.298707, -1.336874, -2.579213, -0.796303, 1.570796, 1.869504],accel_mss,speed_ms,0,blend_radius_m)
  movel([0.299179, -1.336915, -2.579186, -0.796288, 1.570796, 1.869976],accel_mss,speed_ms,0,blend_radius_m)
  movel([0.299654, -1.336970, -2.579150, -0.796269, 1.570796, 1.870450],accel_mss,speed_ms,0,blend_radius_m)
  movel([0.300120, -1.337038, -2.579105, -0.796245, 1.570796, 1.870916],accel_mss,speed_ms,0,blend_radius_m)
  movel([0.300582, -1.337116, -2.579055, -0.796218, 1.570796, 1.871378],accel_mss,speed_ms,0,blend_radius_m)
  movel([0.301004, -1.337201, -2.578999, -0.796189, 1.570796, 1.871800],accel_mss,speed_ms,0,blend_radius_m)
  movel([0.301418, -1.337296, -2.578937, -0.796156, 1.570796, 1.872214],accel_mss,speed_ms,0,blend_radius_m)
  movel([0.301824, -1.337406, -2.578865, -0.796118, 1.570796, 1.872621],accel_mss,speed_ms,0,blend_radius_m)
  movel([0.302367, -1.337574, -2.578756, -0.796059, 1.570796, 1.873163],accel_mss,speed_ms,0,blend_radius_m)
  movel([0.302893, -1.337760, -2.578634, -0.795995, 1.570796, 1.873690],accel_mss,speed_ms,0,blend_radius_m)
  movel([0.303409, -1.337963, -2.578501, -0.795925, 1.570796, 1.874206],accel_mss,speed_ms,0,blend_radius_m)
  movel([0.303912, -1.338184, -2.578357, -0.795848, 1.570796, 1.874708],accel_mss,speed_ms,0,blend_radius_m)
  movel([0.304400, -1.338421, -2.578202, -0.795766, 1.570796, 1.875196],accel_mss,speed_ms,0,blend_radius_m)
  movel([0.304871, -1.338678, -2.578033, -0.795677, 1.570796, 1.875668],accel_mss,speed_ms,0,blend_radius_m)
  movel([0.305329, -1.338949, -2.577856, -0.795584, 1.570796, 1.876125],accel_mss,speed_ms,0,blend_radius_m)
  movel([0.305772, -1.339239, -2.577666, -0.795484, 1.570796, 1.876568],accel_mss,speed_ms,0,blend_radius_m)
  movel([0.306192, -1.339542, -2.577468, -0.795380, 1.570796, 1.876988],accel_mss,speed_ms,0,blend_radius_m)
  movel([0.306597, -1.339860, -2.577259, -0.795270, 1.570796, 1.877393],accel_mss,speed_ms,0,blend_radius_m)
  movel([0.306987, -1.340193, -2.577040, -0.795156, 1.570796, 1.877784],accel_mss,speed_ms,0,blend_radius_m)
  movel([0.307357, -1.340545, -2.576809, -0.795035, 1.570796, 1.878154],accel_mss,speed_ms,0,blend_radius_m)
  movel([0.307710, -1.340910, -2.576569, -0.794910, 1.570796, 1.878507],accel_mss,speed_ms,0,blend_radius_m)
  movel([0.308048, -1.341293, -2.576317, -0.794779, 1.570796, 1.878844],accel_mss,speed_ms,0,blend_radius_m)
  movel([0.308365, -1.341687, -2.576057, -0.794644, 1.570796, 1.879161],accel_mss,speed_ms,0,blend_radius_m)
  movel([0.308666, -1.342099, -2.575786, -0.794504, 1.570796, 1.879462],accel_mss,speed_ms,0,blend_radius_m)
  movel([0.308949, -1.342529, -2.575503, -0.794358, 1.570796, 1.879746],accel_mss,speed_ms,0,blend_radius_m)
  movel([0.309216, -1.342971, -2.575210, -0.794207, 1.570796, 1.880012],accel_mss,speed_ms,0,blend_radius_m)
  movel([0.309464, -1.343428, -2.574909, -0.794053, 1.570796, 1.880260],accel_mss,speed_ms,0,blend_radius_m)
  movel([0.309693, -1.343897, -2.574598, -0.793894, 1.570796, 1.880489],accel_mss,speed_ms,0,blend_radius_m)
  movel([0.309904, -1.344377, -2.574281, -0.793731, 1.570796, 1.880700],accel_mss,speed_ms,0,blend_radius_m)
  movel([0.310093, -1.344871, -2.573953, -0.793565, 1.570796, 1.880890],accel_mss,speed_ms,0,blend_radius_m)
  movel([0.310265, -1.345375, -2.573619, -0.793395, 1.570796, 1.881061],accel_mss,speed_ms,0,blend_radius_m)
  movel([0.310416, -1.345890, -2.573277, -0.793222, 1.570796, 1.881212],accel_mss,speed_ms,0,blend_radius_m)
  movel([0.310553, -1.346434, -2.572915, -0.793040, 1.570796, 1.881349],accel_mss,speed_ms,0,blend_radius_m)
  movel([0.310670, -1.346986, -2.572548, -0.792855, 1.570796, 1.881466],accel_mss,speed_ms,0,blend_radius_m)
  movel([0.310770, -1.347547, -2.572174, -0.792668, 1.570796, 1.881566],accel_mss,speed_ms,0,blend_radius_m)
  movel([0.310852, -1.348118, -2.571793, -0.792478, 1.570796, 1.881649],accel_mss,speed_ms,0,blend_radius_m)
  movel([0.310916, -1.348695, -2.571408, -0.792286, 1.570796, 1.881712],accel_mss,speed_ms,0,blend_radius_m)
  movel([0.310960, -1.349280, -2.571016, -0.792092, 1.570796, 1.881756],accel_mss,speed_ms,0,blend_radius_m)
  movel([0.310984, -1.349874, -2.570619, -0.791896, 1.570796, 1.881781],accel_mss,speed_ms,0,blend_radius_m)
  movel([0.310993, -1.350473, -2.570217, -0.791698, 1.570796, 1.881789],accel_mss,speed_ms,0,blend_radius_m)
  movel([0.310983, -1.350932, -2.569909, -0.791547, 1.570796, 1.881779],accel_mss,speed_ms,0,blend_radius_m)
  movel([0.310955, -1.351395, -2.569598, -0.791395, 1.570796, 1.881751],accel_mss,speed_ms,0,blend_radius_m)
  movel([0.310902, -1.352029, -2.569172, -0.791188, 1.570796, 1.881698],accel_mss,speed_ms,0,blend_radius_m)
  movel([0.310839, -1.352665, -2.568744, -0.790980, 1.570796, 1.881636],accel_mss,speed_ms,0,blend_radius_m)
  movel([0.310771, -1.353291, -2.568322, -0.790776, 1.570796, 1.881567],accel_mss,speed_ms,0,blend_radius_m)
  movel([0.310692, -1.353919, -2.567898, -0.790572, 1.570796, 1.881488],accel_mss,speed_ms,0,blend_radius_m)
  movel([0.310626, -1.354340, -2.567613, -0.790435, 1.570796, 1.881422],accel_mss,speed_ms,0,blend_radius_m)
  movel([0.310542, -1.354766, -2.567325, -0.790297, 1.570796, 1.881338],accel_mss,speed_ms,0,blend_radius_m)
  movel([0.310406, -1.355354, -2.566928, -0.790107, 1.570796, 1.881203],accel_mss,speed_ms,0,blend_radius_m)
  movel([0.310377, -1.355386, -2.566906, -0.790097, 1.570796, 1.881173],accel_mss,speed_ms,0,blend_radius_m)
  movel([0.310335, -1.355415, -2.566886, -0.790088, 1.570796, 1.881131],accel_mss,speed_ms,0,blend_radius_m)
  movel([0.310290, -1.355431, -2.566876, -0.790083, 1.570796, 1.881086],accel_mss,speed_ms,0,blend_radius_m)
  speed_ms = 0.003
  movel([0.310290, -1.358612, -2.568420, -0.785357, 1.570796, 1.881086],accel_mss,speed_ms,0,blend_radius_m)
  speed_ms = 0.007
  movel([0.310214, -1.358629, -2.568408, -0.785352, 1.570796, 1.881011],accel_mss,speed_ms,0,blend_radius_m)
  movel([0.310141, -1.358634, -2.568405, -0.785350, 1.570796, 1.880937],accel_mss,speed_ms,0,blend_radius_m)
  movel([0.309901, -1.358634, -2.568405, -0.785350, 1.570796, 1.880697],accel_mss,speed_ms,0,blend_radius_m)
  movel([0.308940, -1.358622, -2.568413, -0.785354, 1.570796, 1.879736],accel_mss,speed_ms,0,blend_radius_m)
  movel([0.298968, -1.358733, -2.568338, -0.785319, 1.570796, 1.869764],accel_mss,speed_ms,0,blend_radius_m)
  movel([0.288662, -1.358949, -2.568190, -0.785250, 1.570796, 1.859458],accel_mss,speed_ms,0,blend_radius_m)
  movel([0.288310, -1.358976, -2.568172, -0.785241, 1.570796, 1.859107],accel_mss,speed_ms,0,blend_radius_m)
  movel([0.288264, -1.358975, -2.568173, -0.785242, 1.570796, 1.859060],accel_mss,speed_ms,0,blend_radius_m)
  movel([0.288229, -1.358959, -2.568183, -0.785247, 1.570796, 1.859025],accel_mss,speed_ms,0,blend_radius_m)
  movel([0.288203, -1.358929, -2.568204, -0.785256, 1.570796, 1.859000],accel_mss,speed_ms,0,blend_radius_m)
  movel([0.288192, -1.358890, -2.568230, -0.785268, 1.570796, 1.858988],accel_mss,speed_ms,0,blend_radius_m)
  movel([0.288195, -1.358821, -2.568277, -0.785291, 1.570796, 1.858991],accel_mss,speed_ms,0,blend_radius_m)
  movel([0.288208, -1.358751, -2.568325, -0.785313, 1.570796, 1.859004],accel_mss,speed_ms,0,blend_radius_m)
  movel([0.288279, -1.358507, -2.568491, -0.785391, 1.570796, 1.859075],accel_mss,speed_ms,0,blend_radius_m)
  movel([0.288342, -1.358322, -2.568617, -0.785450, 1.570796, 1.859138],accel_mss,speed_ms,0,blend_radius_m)
  movel([0.288415, -1.358133, -2.568746, -0.785511, 1.570796, 1.859211],accel_mss,speed_ms,0,blend_radius_m)
  movel([0.289451, -1.355565, -2.570487, -0.786337, 1.570796, 1.860248],accel_mss,speed_ms,0,blend_radius_m)
  movel([0.290662, -1.352585, -2.572497, -0.787307, 1.570796, 1.861458],accel_mss,speed_ms,0,blend_radius_m)
  movel([0.292076, -1.349129, -2.574812, -0.788448, 1.570796, 1.862872],accel_mss,speed_ms,0,blend_radius_m)
  movel([0.295785, -1.340115, -2.580775, -0.791499, 1.570796, 1.866581],accel_mss,speed_ms,0,blend_radius_m)
  movel([0.296446, -1.340071, -2.580804, -0.791514, 1.570796, 1.867242],accel_mss,speed_ms,0,blend_radius_m)
  movel([0.296887, -1.340046, -2.580820, -0.791522, 1.570796, 1.867683],accel_mss,speed_ms,0,blend_radius_m)
  movel([0.297322, -1.340039, -2.580825, -0.791525, 1.570796, 1.868119],accel_mss,speed_ms,0,blend_radius_m)
  movel([0.297751, -1.340044, -2.580822, -0.791523, 1.570796, 1.868548],accel_mss,speed_ms,0,blend_radius_m)
  movel([0.298232, -1.340065, -2.580808, -0.791516, 1.570796, 1.869029],accel_mss,speed_ms,0,blend_radius_m)
  movel([0.298707, -1.340097, -2.580787, -0.791505, 1.570796, 1.869504],accel_mss,speed_ms,0,blend_radius_m)
  movel([0.299179, -1.340139, -2.580760, -0.791491, 1.570796, 1.869976],accel_mss,speed_ms,0,blend_radius_m)
  movel([0.299654, -1.340194, -2.580724, -0.791472, 1.570796, 1.870450],accel_mss,speed_ms,0,blend_radius_m)
  movel([0.300120, -1.340261, -2.580679, -0.791448, 1.570796, 1.870916],accel_mss,speed_ms,0,blend_radius_m)
  movel([0.300582, -1.340339, -2.580628, -0.791422, 1.570796, 1.871378],accel_mss,speed_ms,0,blend_radius_m)
  movel([0.301004, -1.340424, -2.580573, -0.791392, 1.570796, 1.871800],accel_mss,speed_ms,0,blend_radius_m)
  movel([0.301418, -1.340519, -2.580510, -0.791360, 1.570796, 1.872214],accel_mss,speed_ms,0,blend_radius_m)
  movel([0.301824, -1.340629, -2.580438, -0.791322, 1.570796, 1.872621],accel_mss,speed_ms,0,blend_radius_m)
  movel([0.302367, -1.340796, -2.580329, -0.791264, 1.570796, 1.873163],accel_mss,speed_ms,0,blend_radius_m)
  movel([0.302893, -1.340981, -2.580207, -0.791201, 1.570796, 1.873690],accel_mss,speed_ms,0,blend_radius_m)
  movel([0.303409, -1.341184, -2.580074, -0.791131, 1.570796, 1.874206],accel_mss,speed_ms,0,blend_radius_m)
  movel([0.303912, -1.341405, -2.579929, -0.791055, 1.570796, 1.874708],accel_mss,speed_ms,0,blend_radius_m)
  movel([0.304400, -1.341641, -2.579773, -0.790974, 1.570796, 1.875196],accel_mss,speed_ms,0,blend_radius_m)
  movel([0.304871, -1.341898, -2.579605, -0.790887, 1.570796, 1.875668],accel_mss,speed_ms,0,blend_radius_m)
  movel([0.305329, -1.342168, -2.579427, -0.790794, 1.570796, 1.876125],accel_mss,speed_ms,0,blend_radius_m)
  movel([0.305772, -1.342458, -2.579236, -0.790695, 1.570796, 1.876568],accel_mss,speed_ms,0,blend_radius_m)
  movel([0.306192, -1.342759, -2.579037, -0.790592, 1.570796, 1.876988],accel_mss,speed_ms,0,blend_radius_m)
  movel([0.306597, -1.343077, -2.578828, -0.790484, 1.570796, 1.877393],accel_mss,speed_ms,0,blend_radius_m)
  movel([0.306987, -1.343409, -2.578609, -0.790371, 1.570796, 1.877784],accel_mss,speed_ms,0,blend_radius_m)
  movel([0.307357, -1.343760, -2.578377, -0.790252, 1.570796, 1.878154],accel_mss,speed_ms,0,blend_radius_m)
  movel([0.307710, -1.344125, -2.578136, -0.790128, 1.570796, 1.878507],accel_mss,speed_ms,0,blend_radius_m)
  movel([0.308048, -1.344507, -2.577884, -0.789998, 1.570796, 1.878844],accel_mss,speed_ms,0,blend_radius_m)
  movel([0.308365, -1.344900, -2.577624, -0.789865, 1.570796, 1.879161],accel_mss,speed_ms,0,blend_radius_m)
  movel([0.308666, -1.345311, -2.577352, -0.789726, 1.570796, 1.879462],accel_mss,speed_ms,0,blend_radius_m)
  movel([0.308949, -1.345740, -2.577067, -0.789582, 1.570796, 1.879746],accel_mss,speed_ms,0,blend_radius_m)
  movel([0.309216, -1.346181, -2.576774, -0.789433, 1.570796, 1.880012],accel_mss,speed_ms,0,blend_radius_m)
  movel([0.309464, -1.346636, -2.576472, -0.789280, 1.570796, 1.880260],accel_mss,speed_ms,0,blend_radius_m)
  movel([0.309693, -1.347105, -2.576161, -0.789123, 1.570796, 1.880489],accel_mss,speed_ms,0,blend_radius_m)
  movel([0.309904, -1.347584, -2.575843, -0.788963, 1.570796, 1.880700],accel_mss,speed_ms,0,blend_radius_m)
  movel([0.310093, -1.348076, -2.575515, -0.788798, 1.570796, 1.880890],accel_mss,speed_ms,0,blend_radius_m)
  movel([0.310265, -1.348579, -2.575179, -0.788630, 1.570796, 1.881061],accel_mss,speed_ms,0,blend_radius_m)
  movel([0.310416, -1.349093, -2.574836, -0.788459, 1.570796, 1.881212],accel_mss,speed_ms,0,blend_radius_m)
  movel([0.310553, -1.349636, -2.574474, -0.788279, 1.570796, 1.881349],accel_mss,speed_ms,0,blend_radius_m)
  movel([0.310670, -1.350187, -2.574105, -0.788097, 1.570796, 1.881466],accel_mss,speed_ms,0,blend_radius_m)
  movel([0.310770, -1.350746, -2.573731, -0.787912, 1.570796, 1.881566],accel_mss,speed_ms,0,blend_radius_m)
  movel([0.310852, -1.351316, -2.573349, -0.787724, 1.570796, 1.881649],accel_mss,speed_ms,0,blend_radius_m)
  movel([0.310916, -1.351892, -2.572963, -0.787535, 1.570796, 1.881712],accel_mss,speed_ms,0,blend_radius_m)
  movel([0.310960, -1.352476, -2.572570, -0.787343, 1.570796, 1.881756],accel_mss,speed_ms,0,blend_radius_m)
  movel([0.310984, -1.353068, -2.572172, -0.787149, 1.570796, 1.881781],accel_mss,speed_ms,0,blend_radius_m)
  movel([0.310993, -1.353666, -2.571769, -0.786954, 1.570796, 1.881789],accel_mss,speed_ms,0,blend_radius_m)
  movel([0.310983, -1.354124, -2.571460, -0.786804, 1.570796, 1.881779],accel_mss,speed_ms,0,blend_radius_m)
  movel([0.310955, -1.354586, -2.571149, -0.786654, 1.570796, 1.881751],accel_mss,speed_ms,0,blend_radius_m)
  movel([0.310902, -1.355218, -2.570722, -0.786449, 1.570796, 1.881698],accel_mss,speed_ms,0,blend_radius_m)
  movel([0.310839, -1.355853, -2.570292, -0.786244, 1.570796, 1.881636],accel_mss,speed_ms,0,blend_radius_m)
  movel([0.310771, -1.356477, -2.569870, -0.786042, 1.570796, 1.881567],accel_mss,speed_ms,0,blend_radius_m)
  movel([0.310692, -1.357103, -2.569445, -0.785841, 1.570796, 1.881488],accel_mss,speed_ms,0,blend_radius_m)
  movel([0.310626, -1.357524, -2.569159, -0.785705, 1.570796, 1.881422],accel_mss,speed_ms,0,blend_radius_m)
  movel([0.310542, -1.357949, -2.568870, -0.785569, 1.570796, 1.881338],accel_mss,speed_ms,0,blend_radius_m)
  movel([0.310406, -1.358535, -2.568472, -0.785382, 1.570796, 1.881203],accel_mss,speed_ms,0,blend_radius_m)
  movel([0.310377, -1.358568, -2.568450, -0.785372, 1.570796, 1.881173],accel_mss,speed_ms,0,blend_radius_m)
  movel([0.310335, -1.358596, -2.568430, -0.785362, 1.570796, 1.881131],accel_mss,speed_ms,0,blend_radius_m)
  movel([0.310290, -1.358612, -2.568420, -0.785357, 1.570796, 1.881086],accel_mss,speed_ms,0,blend_radius_m)
  speed_ms = 0.003
  movel([0.310290, -1.346022, -2.562195, -0.804172, 1.570796, 1.881086],accel_mss,speed_ms,0,blend_radius_m)
  speed_ms = 0.01
  movel([0.310290, -1.321918, -2.549368, -0.841103, 1.570796, 1.881086],accel_mss,speed_ms,0,blend_radius_m)
  movel([0.306482, -1.331317, -2.543243, -0.837830, 1.570796, 1.877279],accel_mss,speed_ms,0,blend_radius_m)
  movel([0.306482, -1.355279, -2.555952, -0.801158, 1.570796, 1.877279],accel_mss,speed_ms,0,blend_radius_m)
  speed_ms = 0.003
  movel([0.306482, -1.364626, -2.560588, -0.787175, 1.570796, 1.877279],accel_mss,speed_ms,0,blend_radius_m)
  speed_ms = 0.007
  movel([0.306497, -1.364629, -2.560586, -0.787174, 1.570796, 1.877294],accel_mss,speed_ms,0,blend_radius_m)
  movel([0.306510, -1.364641, -2.560578, -0.787170, 1.570796, 1.877306],accel_mss,speed_ms,0,blend_radius_m)
  movel([0.306504, -1.364664, -2.560562, -0.787163, 1.570796, 1.877301],accel_mss,speed_ms,0,blend_radius_m)
  movel([0.305903, -1.365590, -2.559922, -0.786877, 1.570796, 1.876699],accel_mss,speed_ms,0,blend_radius_m)
  movel([0.305337, -1.366452, -2.559326, -0.786611, 1.570796, 1.876134],accel_mss,speed_ms,0,blend_radius_m)
  movel([0.305113, -1.366783, -2.559096, -0.786510, 1.570796, 1.875909],accel_mss,speed_ms,0,blend_radius_m)
  movel([0.304882, -1.367115, -2.558866, -0.786408, 1.570796, 1.875678],accel_mss,speed_ms,0,blend_radius_m)
  movel([0.304461, -1.367701, -2.558460, -0.786229, 1.570796, 1.875257],accel_mss,speed_ms,0,blend_radius_m)
  movel([0.304026, -1.368281, -2.558056, -0.786052, 1.570796, 1.874822],accel_mss,speed_ms,0,blend_radius_m)
  movel([0.303577, -1.368856, -2.557656, -0.785877, 1.570796, 1.874374],accel_mss,speed_ms,0,blend_radius_m)
  movel([0.303113, -1.369423, -2.557262, -0.785704, 1.570796, 1.873910],accel_mss,speed_ms,0,blend_radius_m)
  movel([0.302640, -1.369984, -2.556870, -0.785535, 1.570796, 1.873436],accel_mss,speed_ms,0,blend_radius_m)
  movel([0.302129, -1.370564, -2.556466, -0.785359, 1.570796, 1.872925],accel_mss,speed_ms,0,blend_radius_m)
  movel([0.301609, -1.371136, -2.556066, -0.785187, 1.570796, 1.872406],accel_mss,speed_ms,0,blend_radius_m)
  movel([0.301079, -1.371699, -2.555672, -0.785018, 1.570796, 1.871875],accel_mss,speed_ms,0,blend_radius_m)
  movel([0.300537, -1.372257, -2.555281, -0.784851, 1.570796, 1.871334],accel_mss,speed_ms,0,blend_radius_m)
  movel([0.299986, -1.372805, -2.554897, -0.784687, 1.570796, 1.870782],accel_mss,speed_ms,0,blend_radius_m)
  movel([0.299427, -1.373342, -2.554520, -0.784527, 1.570796, 1.870223],accel_mss,speed_ms,0,blend_radius_m)
  movel([0.298859, -1.373871, -2.554148, -0.784370, 1.570796, 1.869655],accel_mss,speed_ms,0,blend_radius_m)
  movel([0.298284, -1.374390, -2.553783, -0.784216, 1.570796, 1.869080],accel_mss,speed_ms,0,blend_radius_m)
  movel([0.297698, -1.374901, -2.553423, -0.784064, 1.570796, 1.868494],accel_mss,speed_ms,0,blend_radius_m)
  movel([0.297105, -1.375400, -2.553072, -0.783917, 1.570796, 1.867902],accel_mss,speed_ms,0,blend_radius_m)
  movel([0.296533, -1.375863, -2.552745, -0.783781, 1.570796, 1.867330],accel_mss,speed_ms,0,blend_radius_m)
  movel([0.295956, -1.376317, -2.552425, -0.783648, 1.570796, 1.866752],accel_mss,speed_ms,0,blend_radius_m)
  movel([0.295370, -1.376755, -2.552115, -0.783519, 1.570796, 1.866166],accel_mss,speed_ms,0,blend_radius_m)
  movel([0.294774, -1.377184, -2.551811, -0.783393, 1.570796, 1.865570],accel_mss,speed_ms,0,blend_radius_m)
  movel([0.294174, -1.377599, -2.551518, -0.783272, 1.570796, 1.864970],accel_mss,speed_ms,0,blend_radius_m)
  movel([0.293638, -1.377956, -2.551265, -0.783168, 1.570796, 1.864434],accel_mss,speed_ms,0,blend_radius_m)
  movel([0.293099, -1.378303, -2.551019, -0.783067, 1.570796, 1.863895],accel_mss,speed_ms,0,blend_radius_m)
  movel([0.292554, -1.378640, -2.550780, -0.782969, 1.570796, 1.863350],accel_mss,speed_ms,0,blend_radius_m)
  movel([0.292006, -1.378967, -2.550548, -0.782874, 1.570796, 1.862802],accel_mss,speed_ms,0,blend_radius_m)
  movel([0.291456, -1.379285, -2.550322, -0.782782, 1.570796, 1.862253],accel_mss,speed_ms,0,blend_radius_m)
  movel([0.290901, -1.379593, -2.550103, -0.782693, 1.570796, 1.861697],accel_mss,speed_ms,0,blend_radius_m)
  movel([0.290357, -1.379880, -2.549898, -0.782610, 1.570796, 1.861153],accel_mss,speed_ms,0,blend_radius_m)
  movel([0.289812, -1.380159, -2.549700, -0.782530, 1.570796, 1.860608],accel_mss,speed_ms,0,blend_radius_m)
  movel([0.289261, -1.380426, -2.549510, -0.782453, 1.570796, 1.860057],accel_mss,speed_ms,0,blend_radius_m)
  movel([0.288712, -1.380682, -2.549327, -0.782379, 1.570796, 1.859508],accel_mss,speed_ms,0,blend_radius_m)
  movel([0.288160, -1.380926, -2.549154, -0.782309, 1.570796, 1.858956],accel_mss,speed_ms,0,blend_radius_m)
  movel([0.287607, -1.381159, -2.548988, -0.782243, 1.570796, 1.858404],accel_mss,speed_ms,0,blend_radius_m)
  movel([0.287052, -1.381379, -2.548830, -0.782179, 1.570796, 1.857848],accel_mss,speed_ms,0,blend_radius_m)
  movel([0.286498, -1.381587, -2.548682, -0.782120, 1.570796, 1.857294],accel_mss,speed_ms,0,blend_radius_m)
  movel([0.285944, -1.381782, -2.548543, -0.782064, 1.570796, 1.856740],accel_mss,speed_ms,0,blend_radius_m)
  movel([0.285389, -1.381966, -2.548411, -0.782011, 1.570796, 1.856185],accel_mss,speed_ms,0,blend_radius_m)
  movel([0.284836, -1.382138, -2.548289, -0.781962, 1.570796, 1.855632],accel_mss,speed_ms,0,blend_radius_m)
  movel([0.284284, -1.382297, -2.548175, -0.781917, 1.570796, 1.855081],accel_mss,speed_ms,0,blend_radius_m)
  movel([0.283719, -1.382449, -2.548067, -0.781874, 1.570796, 1.854516],accel_mss,speed_ms,0,blend_radius_m)
  movel([0.283156, -1.382588, -2.547967, -0.781834, 1.570796, 1.853952],accel_mss,speed_ms,0,blend_radius_m)
  movel([0.282595, -1.382714, -2.547877, -0.781798, 1.570796, 1.853391],accel_mss,speed_ms,0,blend_radius_m)
  movel([0.282034, -1.382830, -2.547794, -0.781765, 1.570796, 1.852831],accel_mss,speed_ms,0,blend_radius_m)
  movel([0.281478, -1.382932, -2.547721, -0.781736, 1.570796, 1.852274],accel_mss,speed_ms,0,blend_radius_m)
  movel([0.280924, -1.383022, -2.547656, -0.781711, 1.570796, 1.851720],accel_mss,speed_ms,0,blend_radius_m)
  movel([0.280343, -1.383102, -2.547599, -0.781688, 1.570796, 1.851139],accel_mss,speed_ms,0,blend_radius_m)
  movel([0.279766, -1.383167, -2.547552, -0.781669, 1.570796, 1.850563],accel_mss,speed_ms,0,blend_radius_m)
  movel([0.279126, -1.383225, -2.547511, -0.781653, 1.570796, 1.849923],accel_mss,speed_ms,0,blend_radius_m)
  movel([0.278493, -1.383270, -2.547479, -0.781640, 1.570796, 1.849289],accel_mss,speed_ms,0,blend_radius_m)
  movel([0.277894, -1.383302, -2.547455, -0.781631, 1.570796, 1.848691],accel_mss,speed_ms,0,blend_radius_m)
  movel([0.277297, -1.383333, -2.547434, -0.781622, 1.570796, 1.848093],accel_mss,speed_ms,0,blend_radius_m)
  movel([0.277230, -1.383328, -2.547437, -0.781624, 1.570796, 1.848027],accel_mss,speed_ms,0,blend_radius_m)
  movel([0.277171, -1.383314, -2.547447, -0.781628, 1.570796, 1.847967],accel_mss,speed_ms,0,blend_radius_m)
  movel([0.277120, -1.383288, -2.547466, -0.781635, 1.570796, 1.847916],accel_mss,speed_ms,0,blend_radius_m)
  movel([0.277078, -1.383252, -2.547491, -0.781645, 1.570796, 1.847875],accel_mss,speed_ms,0,blend_radius_m)
  movel([0.277063, -1.383226, -2.547510, -0.781653, 1.570796, 1.847860],accel_mss,speed_ms,0,blend_radius_m)
  movel([0.277062, -1.383194, -2.547533, -0.781662, 1.570796, 1.847858],accel_mss,speed_ms,0,blend_radius_m)
  movel([0.277071, -1.383157, -2.547560, -0.781672, 1.570796, 1.847867],accel_mss,speed_ms,0,blend_radius_m)
  movel([0.280441, -1.374678, -2.553580, -0.784130, 1.570796, 1.851237],accel_mss,speed_ms,0,blend_radius_m)
  movel([0.283691, -1.366559, -2.559251, -0.786579, 1.570796, 1.854487],accel_mss,speed_ms,0,blend_radius_m)
  movel([0.283849, -1.366172, -2.559519, -0.786698, 1.570796, 1.854646],accel_mss,speed_ms,0,blend_radius_m)
  movel([0.284019, -1.365786, -2.559787, -0.786817, 1.570796, 1.854816],accel_mss,speed_ms,0,blend_radius_m)
  movel([0.284199, -1.365398, -2.560055, -0.786936, 1.570796, 1.854995],accel_mss,speed_ms,0,blend_radius_m)
  movel([0.284422, -1.364928, -2.560380, -0.787082, 1.570796, 1.855219],accel_mss,speed_ms,0,blend_radius_m)
  movel([0.295474, -1.364717, -2.560525, -0.787147, 1.570796, 1.866271],accel_mss,speed_ms,0,blend_radius_m)
  movel([0.299702, -1.364666, -2.560560, -0.787162, 1.570796, 1.870498],accel_mss,speed_ms,0,blend_radius_m)
  movel([0.303258, -1.364640, -2.560578, -0.787171, 1.570796, 1.874055],accel_mss,speed_ms,0,blend_radius_m)
  movel([0.306482, -1.364626, -2.560588, -0.787175, 1.570796, 1.877279],accel_mss,speed_ms,0,blend_radius_m)
  speed_ms = 0.003
  movel([0.306482, -1.367786, -2.562117, -0.782486, 1.570796, 1.877279],accel_mss,speed_ms,0,blend_radius_m)
  speed_ms = 0.007
  movel([0.306497, -1.367789, -2.562115, -0.782485, 1.570796, 1.877294],accel_mss,speed_ms,0,blend_radius_m)
  movel([0.306510, -1.367801, -2.562107, -0.782481, 1.570796, 1.877306],accel_mss,speed_ms,0,blend_radius_m)
  movel([0.306504, -1.367824, -2.562091, -0.782474, 1.570796, 1.877301],accel_mss,speed_ms,0,blend_radius_m)
  movel([0.305903, -1.368748, -2.561450, -0.782192, 1.570796, 1.876699],accel_mss,speed_ms,0,blend_radius_m)
  movel([0.305337, -1.369608, -2.560852, -0.781930, 1.570796, 1.876134],accel_mss,speed_ms,0,blend_radius_m)
  movel([0.305113, -1.369938, -2.560622, -0.781829, 1.570796, 1.875909],accel_mss,speed_ms,0,blend_radius_m)
  movel([0.304882, -1.370269, -2.560391, -0.781729, 1.570796, 1.875678],accel_mss,speed_ms,0,blend_radius_m)
  movel([0.304461, -1.370853, -2.559984, -0.781552, 1.570796, 1.875257],accel_mss,speed_ms,0,blend_radius_m)
  movel([0.304026, -1.371432, -2.559580, -0.781377, 1.570796, 1.874822],accel_mss,speed_ms,0,blend_radius_m)
  movel([0.303577, -1.372006, -2.559179, -0.781204, 1.570796, 1.874374],accel_mss,speed_ms,0,blend_radius_m)
  movel([0.303113, -1.372572, -2.558783, -0.781034, 1.570796, 1.873910],accel_mss,speed_ms,0,blend_radius_m)
  movel([0.302640, -1.373131, -2.558391, -0.780867, 1.570796, 1.873436],accel_mss,speed_ms,0,blend_radius_m)
  movel([0.302129, -1.373710, -2.557985, -0.780694, 1.570796, 1.872925],accel_mss,speed_ms,0,blend_radius_m)
  movel([0.301609, -1.374280, -2.557585, -0.780524, 1.570796, 1.872406],accel_mss,speed_ms,0,blend_radius_m)
  movel([0.301079, -1.374843, -2.557189, -0.780357, 1.570796, 1.871875],accel_mss,speed_ms,0,blend_radius_m)
  movel([0.300537, -1.375399, -2.556798, -0.780192, 1.570796, 1.871334],accel_mss,speed_ms,0,blend_radius_m)
  movel([0.299986, -1.375946, -2.556413, -0.780031, 1.570796, 1.870782],accel_mss,speed_ms,0,blend_radius_m)
  movel([0.299427, -1.376482, -2.556035, -0.779873, 1.570796, 1.870223],accel_mss,speed_ms,0,blend_radius_m)
  movel([0.298859, -1.377009, -2.555662, -0.779717, 1.570796, 1.869655],accel_mss,speed_ms,0,blend_radius_m)
  movel([0.298284, -1.377527, -2.555296, -0.779565, 1.570796, 1.869080],accel_mss,speed_ms,0,blend_radius_m)
  movel([0.297698, -1.378037, -2.554936, -0.779416, 1.570796, 1.868494],accel_mss,speed_ms,0,blend_radius_m)
  movel([0.297105, -1.378534, -2.554584, -0.779271, 1.570796, 1.867902],accel_mss,speed_ms,0,blend_radius_m)
  movel([0.296533, -1.378997, -2.554256, -0.779136, 1.570796, 1.867330],accel_mss,speed_ms,0,blend_radius_m)
  movel([0.295956, -1.379449, -2.553935, -0.779005, 1.570796, 1.866752],accel_mss,speed_ms,0,blend_radius_m)
  movel([0.295370, -1.379886, -2.553624, -0.778878, 1.570796, 1.866166],accel_mss,speed_ms,0,blend_radius_m)
  movel([0.294774, -1.380314, -2.553320, -0.778754, 1.570796, 1.865570],accel_mss,speed_ms,0,blend_radius_m)
  movel([0.294174, -1.380728, -2.553026, -0.778635, 1.570796, 1.864970],accel_mss,speed_ms,0,blend_radius_m)
  movel([0.293638, -1.381084, -2.552772, -0.778532, 1.570796, 1.864434],accel_mss,speed_ms,0,blend_radius_m)
  movel([0.293099, -1.381431, -2.552526, -0.778433, 1.570796, 1.863895],accel_mss,speed_ms,0,blend_radius_m)
  movel([0.292554, -1.381767, -2.552286, -0.778336, 1.570796, 1.863350],accel_mss,speed_ms,0,blend_radius_m)
  movel([0.292006, -1.382092, -2.552054, -0.778243, 1.570796, 1.862802],accel_mss,speed_ms,0,blend_radius_m)
  movel([0.291456, -1.382410, -2.551827, -0.778152, 1.570796, 1.862253],accel_mss,speed_ms,0,blend_radius_m)
  movel([0.290901, -1.382717, -2.551608, -0.778064, 1.570796, 1.861697],accel_mss,speed_ms,0,blend_radius_m)
  movel([0.290357, -1.383004, -2.551403, -0.777982, 1.570796, 1.861153],accel_mss,speed_ms,0,blend_radius_m)
  movel([0.289812, -1.383282, -2.551204, -0.777903, 1.570796, 1.860608],accel_mss,speed_ms,0,blend_radius_m)
  movel([0.289261, -1.383548, -2.551014, -0.777827, 1.570796, 1.860057],accel_mss,speed_ms,0,blend_radius_m)
  movel([0.288712, -1.383804, -2.550831, -0.777755, 1.570796, 1.859508],accel_mss,speed_ms,0,blend_radius_m)
  movel([0.288160, -1.384046, -2.550657, -0.777686, 1.570796, 1.858956],accel_mss,speed_ms,0,blend_radius_m)
  movel([0.287607, -1.384279, -2.550490, -0.777620, 1.570796, 1.858404],accel_mss,speed_ms,0,blend_radius_m)
  movel([0.287052, -1.384499, -2.550333, -0.777557, 1.570796, 1.857848],accel_mss,speed_ms,0,blend_radius_m)
  movel([0.286498, -1.384706, -2.550184, -0.777499, 1.570796, 1.857294],accel_mss,speed_ms,0,blend_radius_m)
  movel([0.285944, -1.384901, -2.550045, -0.777444, 1.570796, 1.856740],accel_mss,speed_ms,0,blend_radius_m)
  movel([0.285389, -1.385085, -2.549913, -0.777392, 1.570796, 1.856185],accel_mss,speed_ms,0,blend_radius_m)
  movel([0.284836, -1.385256, -2.549790, -0.777344, 1.570796, 1.855632],accel_mss,speed_ms,0,blend_radius_m)
  movel([0.284284, -1.385414, -2.549676, -0.777299, 1.570796, 1.855081],accel_mss,speed_ms,0,blend_radius_m)
  movel([0.283719, -1.385566, -2.549567, -0.777256, 1.570796, 1.854516],accel_mss,speed_ms,0,blend_radius_m)
  movel([0.283156, -1.385704, -2.549467, -0.777217, 1.570796, 1.853952],accel_mss,speed_ms,0,blend_radius_m)
  movel([0.282595, -1.385830, -2.549377, -0.777182, 1.570796, 1.853391],accel_mss,speed_ms,0,blend_radius_m)
  movel([0.282034, -1.385946, -2.549294, -0.777149, 1.570796, 1.852831],accel_mss,speed_ms,0,blend_radius_m)
  movel([0.281478, -1.386048, -2.549220, -0.777120, 1.570796, 1.852274],accel_mss,speed_ms,0,blend_radius_m)
  movel([0.280924, -1.386138, -2.549156, -0.777095, 1.570796, 1.851720],accel_mss,speed_ms,0,blend_radius_m)
  movel([0.280343, -1.386218, -2.549098, -0.777073, 1.570796, 1.851139],accel_mss,speed_ms,0,blend_radius_m)
  movel([0.279766, -1.386283, -2.549051, -0.777055, 1.570796, 1.850563],accel_mss,speed_ms,0,blend_radius_m)
  movel([0.279126, -1.386341, -2.549010, -0.777038, 1.570796, 1.849923],accel_mss,speed_ms,0,blend_radius_m)
  movel([0.278493, -1.386385, -2.548978, -0.777026, 1.570796, 1.849289],accel_mss,speed_ms,0,blend_radius_m)
  movel([0.277894, -1.386418, -2.548955, -0.777017, 1.570796, 1.848691],accel_mss,speed_ms,0,blend_radius_m)
  movel([0.277297, -1.386448, -2.548933, -0.777008, 1.570796, 1.848093],accel_mss,speed_ms,0,blend_radius_m)
  movel([0.277230, -1.386443, -2.548936, -0.777010, 1.570796, 1.848027],accel_mss,speed_ms,0,blend_radius_m)
  movel([0.277171, -1.386429, -2.548947, -0.777014, 1.570796, 1.847967],accel_mss,speed_ms,0,blend_radius_m)
  movel([0.277120, -1.386403, -2.548965, -0.777021, 1.570796, 1.847916],accel_mss,speed_ms,0,blend_radius_m)
  movel([0.277078, -1.386367, -2.548991, -0.777031, 1.570796, 1.847875],accel_mss,speed_ms,0,blend_radius_m)
  movel([0.277063, -1.386341, -2.549009, -0.777038, 1.570796, 1.847860],accel_mss,speed_ms,0,blend_radius_m)
  movel([0.277062, -1.386310, -2.549032, -0.777047, 1.570796, 1.847858],accel_mss,speed_ms,0,blend_radius_m)
  movel([0.277071, -1.386272, -2.549059, -0.777058, 1.570796, 1.847867],accel_mss,speed_ms,0,blend_radius_m)
  movel([0.280441, -1.377814, -2.555093, -0.779481, 1.570796, 1.851237],accel_mss,speed_ms,0,blend_radius_m)
  movel([0.283691, -1.369714, -2.560777, -0.781897, 1.570796, 1.854487],accel_mss,speed_ms,0,blend_radius_m)
  movel([0.283849, -1.369328, -2.561046, -0.782015, 1.570796, 1.854646],accel_mss,speed_ms,0,blend_radius_m)
  movel([0.284019, -1.368943, -2.561314, -0.782132, 1.570796, 1.854816],accel_mss,speed_ms,0,blend_radius_m)
  movel([0.284199, -1.368556, -2.561583, -0.782250, 1.570796, 1.854995],accel_mss,speed_ms,0,blend_radius_m)
  movel([0.284422, -1.368087, -2.561908, -0.782394, 1.570796, 1.855219],accel_mss,speed_ms,0,blend_radius_m)
  movel([0.295474, -1.367877, -2.562054, -0.782458, 1.570796, 1.866271],accel_mss,speed_ms,0,blend_radius_m)
  movel([0.299702, -1.367826, -2.562089, -0.782473, 1.570796, 1.870498],accel_mss,speed_ms,0,blend_radius_m)
  movel([0.303258, -1.367800, -2.562107, -0.782482, 1.570796, 1.874055],accel_mss,speed_ms,0,blend_radius_m)
  movel([0.306482, -1.367786, -2.562117, -0.782486, 1.570796, 1.877279],accel_mss,speed_ms,0,blend_radius_m)
  speed_ms = 0.003
  movel([0.306482, -1.355279, -2.555952, -0.801158, 1.570796, 1.877279],accel_mss,speed_ms,0,blend_radius_m)
  speed_ms = 0.01
  movel([0.306482, -1.331317, -2.543243, -0.837830, 1.570796, 1.877279],accel_mss,speed_ms,0,blend_radius_m)
  movel([0.281967, -1.366505, -2.519283, -0.826601, 1.570796, 1.852763],accel_mss,speed_ms,0,blend_radius_m)
  movel([0.281967, -1.389907, -2.531555, -0.790927, 1.570796, 1.852763],accel_mss,speed_ms,0,blend_radius_m)
  speed_ms = 0.003
  movel([0.281967, -1.399014, -2.536026, -0.777349, 1.570796, 1.852763],accel_mss,speed_ms,0,blend_radius_m)
  speed_ms = 0.007
  movel([0.282101, -1.399065, -2.535989, -0.777336, 1.570796, 1.852897],accel_mss,speed_ms,0,blend_radius_m)
  movel([0.282114, -1.399078, -2.535979, -0.777332, 1.570796, 1.852911],accel_mss,speed_ms,0,blend_radius_m)
  movel([0.282112, -1.399099, -2.535963, -0.777327, 1.570796, 1.852909],accel_mss,speed_ms,0,blend_radius_m)
  movel([0.282087, -1.399160, -2.535918, -0.777311, 1.570796, 1.852883],accel_mss,speed_ms,0,blend_radius_m)
  movel([0.281403, -1.400355, -2.535034, -0.777000, 1.570796, 1.852199],accel_mss,speed_ms,0,blend_radius_m)
  movel([0.280637, -1.401693, -2.534042, -0.776654, 1.570796, 1.851433],accel_mss,speed_ms,0,blend_radius_m)
  movel([0.279737, -1.403261, -2.532876, -0.776252, 1.570796, 1.850533],accel_mss,speed_ms,0,blend_radius_m)
  movel([0.278835, -1.404826, -2.531708, -0.775855, 1.570796, 1.849631],accel_mss,speed_ms,0,blend_radius_m)
  movel([0.278067, -1.406147, -2.530720, -0.775522, 1.570796, 1.848863],accel_mss,speed_ms,0,blend_radius_m)
  movel([0.277379, -1.407328, -2.529835, -0.775226, 1.570796, 1.848176],accel_mss,speed_ms,0,blend_radius_m)
  movel([0.277360, -1.407354, -2.529815, -0.775220, 1.570796, 1.848156],accel_mss,speed_ms,0,blend_radius_m)
  movel([0.277335, -1.407378, -2.529797, -0.775214, 1.570796, 1.848131],accel_mss,speed_ms,0,blend_radius_m)
  movel([0.277311, -1.407391, -2.529788, -0.775211, 1.570796, 1.848108],accel_mss,speed_ms,0,blend_radius_m)
  movel([0.277285, -1.407396, -2.529784, -0.775209, 1.570796, 1.848082],accel_mss,speed_ms,0,blend_radius_m)
  movel([0.276947, -1.407366, -2.529806, -0.775217, 1.570796, 1.847743],accel_mss,speed_ms,0,blend_radius_m)
  movel([0.276557, -1.407324, -2.529838, -0.775227, 1.570796, 1.847353],accel_mss,speed_ms,0,blend_radius_m)
  movel([0.276107, -1.407266, -2.529881, -0.775242, 1.570796, 1.846903],accel_mss,speed_ms,0,blend_radius_m)
  movel([0.268401, -1.406335, -2.530579, -0.775474, 1.570796, 1.839198],accel_mss,speed_ms,0,blend_radius_m)
  movel([0.266203, -1.406068, -2.530779, -0.775541, 1.570796, 1.836999],accel_mss,speed_ms,0,blend_radius_m)
  movel([0.265171, -1.405938, -2.530877, -0.775574, 1.570796, 1.835967],accel_mss,speed_ms,0,blend_radius_m)
  movel([0.264146, -1.405795, -2.530984, -0.775610, 1.570796, 1.834942],accel_mss,speed_ms,0,blend_radius_m)
  movel([0.263129, -1.405642, -2.531098, -0.775649, 1.570796, 1.833925],accel_mss,speed_ms,0,blend_radius_m)
  movel([0.262318, -1.405510, -2.531197, -0.775682, 1.570796, 1.833114],accel_mss,speed_ms,0,blend_radius_m)
  movel([0.261517, -1.405365, -2.531306, -0.775718, 1.570796, 1.832314],accel_mss,speed_ms,0,blend_radius_m)
  movel([0.260722, -1.405208, -2.531423, -0.775758, 1.570796, 1.831518],accel_mss,speed_ms,0,blend_radius_m)
  movel([0.259973, -1.405049, -2.531542, -0.775798, 1.570796, 1.830770],accel_mss,speed_ms,0,blend_radius_m)
  movel([0.259236, -1.404875, -2.531672, -0.775842, 1.570796, 1.830032],accel_mss,speed_ms,0,blend_radius_m)
  movel([0.258506, -1.404689, -2.531811, -0.775889, 1.570796, 1.829302],accel_mss,speed_ms,0,blend_radius_m)
  movel([0.257924, -1.404525, -2.531933, -0.775931, 1.570796, 1.828721],accel_mss,speed_ms,0,blend_radius_m)
  movel([0.257349, -1.404349, -2.532065, -0.775975, 1.570796, 1.828145],accel_mss,speed_ms,0,blend_radius_m)
  movel([0.256786, -1.404158, -2.532207, -0.776024, 1.570796, 1.827582],accel_mss,speed_ms,0,blend_radius_m)
  movel([0.256230, -1.403957, -2.532357, -0.776075, 1.570796, 1.827027],accel_mss,speed_ms,0,blend_radius_m)
  movel([0.255685, -1.403743, -2.532517, -0.776129, 1.570796, 1.826481],accel_mss,speed_ms,0,blend_radius_m)
  movel([0.255307, -1.403579, -2.532639, -0.776171, 1.570796, 1.826104],accel_mss,speed_ms,0,blend_radius_m)
  movel([0.254940, -1.403404, -2.532770, -0.776216, 1.570796, 1.825736],accel_mss,speed_ms,0,blend_radius_m)
  movel([0.254584, -1.403216, -2.532909, -0.776264, 1.570796, 1.825380],accel_mss,speed_ms,0,blend_radius_m)
  movel([0.254236, -1.403018, -2.533057, -0.776314, 1.570796, 1.825032],accel_mss,speed_ms,0,blend_radius_m)
  movel([0.253901, -1.402806, -2.533215, -0.776368, 1.570796, 1.824697],accel_mss,speed_ms,0,blend_radius_m)
  movel([0.253577, -1.402582, -2.533381, -0.776426, 1.570796, 1.824374],accel_mss,speed_ms,0,blend_radius_m)
  movel([0.253308, -1.402380, -2.533532, -0.776478, 1.570796, 1.824104],accel_mss,speed_ms,0,blend_radius_m)
  movel([0.253051, -1.402163, -2.533693, -0.776533, 1.570796, 1.823847],accel_mss,speed_ms,0,blend_radius_m)
  movel([0.252808, -1.401937, -2.533861, -0.776591, 1.570796, 1.823605],accel_mss,speed_ms,0,blend_radius_m)
  movel([0.252575, -1.401699, -2.534038, -0.776653, 1.570796, 1.823372],accel_mss,speed_ms,0,blend_radius_m)
  movel([0.252356, -1.401451, -2.534222, -0.776717, 1.570796, 1.823152],accel_mss,speed_ms,0,blend_radius_m)
  movel([0.252151, -1.401192, -2.534413, -0.776783, 1.570796, 1.822947],accel_mss,speed_ms,0,blend_radius_m)
  movel([0.251980, -1.400946, -2.534596, -0.776847, 1.570796, 1.822776],accel_mss,speed_ms,0,blend_radius_m)
  movel([0.251825, -1.400689, -2.534787, -0.776913, 1.570796, 1.822622],accel_mss,speed_ms,0,blend_radius_m)
  movel([0.251690, -1.400419, -2.534987, -0.776983, 1.570796, 1.822486],accel_mss,speed_ms,0,blend_radius_m)
  movel([0.251571, -1.400139, -2.535194, -0.777056, 1.570796, 1.822367],accel_mss,speed_ms,0,blend_radius_m)
  movel([0.251468, -1.399848, -2.535410, -0.777132, 1.570796, 1.822264],accel_mss,speed_ms,0,blend_radius_m)
  movel([0.251385, -1.399548, -2.535632, -0.777210, 1.570796, 1.822182],accel_mss,speed_ms,0,blend_radius_m)
  movel([0.251326, -1.399278, -2.535831, -0.777280, 1.570796, 1.822122],accel_mss,speed_ms,0,blend_radius_m)
  movel([0.251281, -1.399003, -2.536034, -0.777352, 1.570796, 1.822077],accel_mss,speed_ms,0,blend_radius_m)
  movel([0.251247, -1.398721, -2.536242, -0.777426, 1.570796, 1.822043],accel_mss,speed_ms,0,blend_radius_m)
  movel([0.251229, -1.398470, -2.536427, -0.777491, 1.570796, 1.822025],accel_mss,speed_ms,0,blend_radius_m)
  movel([0.251228, -1.398213, -2.536617, -0.777559, 1.570796, 1.822025],accel_mss,speed_ms,0,blend_radius_m)
  movel([0.251243, -1.397951, -2.536811, -0.777628, 1.570796, 1.822039],accel_mss,speed_ms,0,blend_radius_m)
  movel([0.251276, -1.397661, -2.537024, -0.777704, 1.570796, 1.822072],accel_mss,speed_ms,0,blend_radius_m)
  movel([0.251323, -1.397370, -2.537239, -0.777781, 1.570796, 1.822119],accel_mss,speed_ms,0,blend_radius_m)
  movel([0.251384, -1.397076, -2.537455, -0.777858, 1.570796, 1.822180],accel_mss,speed_ms,0,blend_radius_m)
  movel([0.251482, -1.396690, -2.537739, -0.777960, 1.570796, 1.822278],accel_mss,speed_ms,0,blend_radius_m)
  movel([0.251585, -1.396303, -2.538023, -0.778063, 1.570796, 1.822381],accel_mss,speed_ms,0,blend_radius_m)
  movel([0.251699, -1.395917, -2.538307, -0.778165, 1.570796, 1.822495],accel_mss,speed_ms,0,blend_radius_m)
  movel([0.251879, -1.395339, -2.538731, -0.778319, 1.570796, 1.822675],accel_mss,speed_ms,0,blend_radius_m)
  movel([0.252046, -1.394842, -2.539095, -0.778452, 1.570796, 1.822842],accel_mss,speed_ms,0,blend_radius_m)
  movel([0.252194, -1.394415, -2.539408, -0.778566, 1.570796, 1.822991],accel_mss,speed_ms,0,blend_radius_m)
  movel([0.252213, -1.394381, -2.539433, -0.778575, 1.570796, 1.823009],accel_mss,speed_ms,0,blend_radius_m)
  movel([0.252239, -1.394352, -2.539454, -0.778583, 1.570796, 1.823035],accel_mss,speed_ms,0,blend_radius_m)
  movel([0.252263, -1.394338, -2.539464, -0.778587, 1.570796, 1.823059],accel_mss,speed_ms,0,blend_radius_m)
  movel([0.252288, -1.394329, -2.539471, -0.778589, 1.570796, 1.823084],accel_mss,speed_ms,0,blend_radius_m)
  movel([0.252311, -1.394328, -2.539472, -0.778589, 1.570796, 1.823107],accel_mss,speed_ms,0,blend_radius_m)
  movel([0.256557, -1.394912, -2.539044, -0.778433, 1.570796, 1.827354],accel_mss,speed_ms,0,blend_radius_m)
  movel([0.261236, -1.395592, -2.538545, -0.778252, 1.570796, 1.832032],accel_mss,speed_ms,0,blend_radius_m)
  movel([0.266759, -1.396441, -2.537922, -0.778026, 1.570796, 1.837555],accel_mss,speed_ms,0,blend_radius_m)
  movel([0.272287, -1.397335, -2.537264, -0.777790, 1.570796, 1.843084],accel_mss,speed_ms,0,blend_radius_m)
  movel([0.277015, -1.398131, -2.536678, -0.777580, 1.570796, 1.847812],accel_mss,speed_ms,0,blend_radius_m)
  movel([0.281147, -1.398847, -2.536149, -0.777393, 1.570796, 1.851943],accel_mss,speed_ms,0,blend_radius_m)
  movel([0.281794, -1.398966, -2.536062, -0.777362, 1.570796, 1.852590],accel_mss,speed_ms,0,blend_radius_m)
  movel([0.281967, -1.399014, -2.536026, -0.777349, 1.570796, 1.852763],accel_mss,speed_ms,0,blend_radius_m)
  speed_ms = 0.003
  movel([0.281967, -1.402090, -2.537500, -0.772799, 1.570796, 1.852763],accel_mss,speed_ms,0,blend_radius_m)
  speed_ms = 0.007
  movel([0.282101, -1.402141, -2.537463, -0.772786, 1.570796, 1.852897],accel_mss,speed_ms,0,blend_radius_m)
  movel([0.282114, -1.402154, -2.537453, -0.772782, 1.570796, 1.852911],accel_mss,speed_ms,0,blend_radius_m)
  movel([0.282112, -1.402175, -2.537437, -0.772777, 1.570796, 1.852909],accel_mss,speed_ms,0,blend_radius_m)
  movel([0.282087, -1.402236, -2.537392, -0.772761, 1.570796, 1.852883],accel_mss,speed_ms,0,blend_radius_m)
  movel([0.281403, -1.403428, -2.536506, -0.772455, 1.570796, 1.852199],accel_mss,speed_ms,0,blend_radius_m)
  movel([0.280637, -1.404762, -2.535512, -0.772115, 1.570796, 1.851433],accel_mss,speed_ms,0,blend_radius_m)
  movel([0.279737, -1.406327, -2.534343, -0.771719, 1.570796, 1.850533],accel_mss,speed_ms,0,blend_radius_m)
  movel([0.278835, -1.407888, -2.533173, -0.771328, 1.570796, 1.849631],accel_mss,speed_ms,0,blend_radius_m)
  movel([0.278067, -1.409206, -2.532183, -0.771000, 1.570796, 1.848863],accel_mss,speed_ms,0,blend_radius_m)
  movel([0.277379, -1.410383, -2.531296, -0.770710, 1.570796, 1.848176],accel_mss,speed_ms,0,blend_radius_m)
  movel([0.277360, -1.410410, -2.531276, -0.770703, 1.570796, 1.848156],accel_mss,speed_ms,0,blend_radius_m)
  movel([0.277335, -1.410433, -2.531258, -0.770698, 1.570796, 1.848131],accel_mss,speed_ms,0,blend_radius_m)
  movel([0.277311, -1.410446, -2.531249, -0.770694, 1.570796, 1.848108],accel_mss,speed_ms,0,blend_radius_m)
  movel([0.277285, -1.410451, -2.531245, -0.770693, 1.570796, 1.848082],accel_mss,speed_ms,0,blend_radius_m)
  movel([0.276947, -1.410421, -2.531267, -0.770700, 1.570796, 1.847743],accel_mss,speed_ms,0,blend_radius_m)
  movel([0.276557, -1.410379, -2.531299, -0.770711, 1.570796, 1.847353],accel_mss,speed_ms,0,blend_radius_m)
  movel([0.276107, -1.410321, -2.531343, -0.770725, 1.570796, 1.846903],accel_mss,speed_ms,0,blend_radius_m)
  movel([0.268401, -1.409393, -2.532042, -0.770954, 1.570796, 1.839198],accel_mss,speed_ms,0,blend_radius_m)
  movel([0.266203, -1.409127, -2.532242, -0.771020, 1.570796, 1.836999],accel_mss,speed_ms,0,blend_radius_m)
  movel([0.265171, -1.408996, -2.532340, -0.771052, 1.570796, 1.835967],accel_mss,speed_ms,0,blend_radius_m)
  movel([0.264146, -1.408854, -2.532448, -0.771088, 1.570796, 1.834942],accel_mss,speed_ms,0,blend_radius_m)
  movel([0.263129, -1.408701, -2.532562, -0.771125, 1.570796, 1.833925],accel_mss,speed_ms,0,blend_radius_m)
  movel([0.262318, -1.408570, -2.532661, -0.771158, 1.570796, 1.833114],accel_mss,speed_ms,0,blend_radius_m)
  movel([0.261517, -1.408425, -2.532770, -0.771194, 1.570796, 1.832314],accel_mss,speed_ms,0,blend_radius_m)
  movel([0.260722, -1.408268, -2.532888, -0.771233, 1.570796, 1.831518],accel_mss,speed_ms,0,blend_radius_m)
  movel([0.259973, -1.408110, -2.533006, -0.771272, 1.570796, 1.830770],accel_mss,speed_ms,0,blend_radius_m)
  movel([0.259236, -1.407937, -2.533137, -0.771316, 1.570796, 1.830032],accel_mss,speed_ms,0,blend_radius_m)
  movel([0.258506, -1.407751, -2.533276, -0.771362, 1.570796, 1.829302],accel_mss,speed_ms,0,blend_radius_m)
  movel([0.257924, -1.407587, -2.533399, -0.771403, 1.570796, 1.828721],accel_mss,speed_ms,0,blend_radius_m)
  movel([0.257349, -1.407411, -2.533531, -0.771447, 1.570796, 1.828145],accel_mss,speed_ms,0,blend_radius_m)
  movel([0.256786, -1.407222, -2.533673, -0.771494, 1.570796, 1.827582],accel_mss,speed_ms,0,blend_radius_m)
  movel([0.256230, -1.407021, -2.533823, -0.771545, 1.570796, 1.827027],accel_mss,speed_ms,0,blend_radius_m)
  movel([0.255685, -1.406807, -2.533984, -0.771598, 1.570796, 1.826481],accel_mss,speed_ms,0,blend_radius_m)
  movel([0.255307, -1.406644, -2.534106, -0.771639, 1.570796, 1.826104],accel_mss,speed_ms,0,blend_radius_m)
  movel([0.254940, -1.406469, -2.534237, -0.771683, 1.570796, 1.825736],accel_mss,speed_ms,0,blend_radius_m)
  movel([0.254584, -1.406282, -2.534377, -0.771730, 1.570796, 1.825380],accel_mss,speed_ms,0,blend_radius_m)
  movel([0.254236, -1.406084, -2.534525, -0.771780, 1.570796, 1.825032],accel_mss,speed_ms,0,blend_radius_m)
  movel([0.253901, -1.405873, -2.534683, -0.771834, 1.570796, 1.824697],accel_mss,speed_ms,0,blend_radius_m)
  movel([0.253577, -1.405649, -2.534850, -0.771890, 1.570796, 1.824374],accel_mss,speed_ms,0,blend_radius_m)
  movel([0.253308, -1.405447, -2.535001, -0.771941, 1.570796, 1.824104],accel_mss,speed_ms,0,blend_radius_m)
  movel([0.253051, -1.405231, -2.535162, -0.771996, 1.570796, 1.823847],accel_mss,speed_ms,0,blend_radius_m)
  movel([0.252808, -1.405006, -2.535330, -0.772053, 1.570796, 1.823605],accel_mss,speed_ms,0,blend_radius_m)
  movel([0.252575, -1.404768, -2.535508, -0.772113, 1.570796, 1.823372],accel_mss,speed_ms,0,blend_radius_m)
  movel([0.252356, -1.404521, -2.535692, -0.772176, 1.570796, 1.823152],accel_mss,speed_ms,0,blend_radius_m)
  movel([0.252151, -1.404263, -2.535884, -0.772242, 1.570796, 1.822947],accel_mss,speed_ms,0,blend_radius_m)
  movel([0.251980, -1.404017, -2.536067, -0.772304, 1.570796, 1.822776],accel_mss,speed_ms,0,blend_radius_m)
  movel([0.251825, -1.403761, -2.536258, -0.772370, 1.570796, 1.822622],accel_mss,speed_ms,0,blend_radius_m)
  movel([0.251690, -1.403492, -2.536459, -0.772439, 1.570796, 1.822486],accel_mss,speed_ms,0,blend_radius_m)
  movel([0.251571, -1.403212, -2.536667, -0.772510, 1.570796, 1.822367],accel_mss,speed_ms,0,blend_radius_m)
  movel([0.251468, -1.402922, -2.536883, -0.772585, 1.570796, 1.822264],accel_mss,speed_ms,0,blend_radius_m)
  movel([0.251385, -1.402622, -2.537105, -0.772662, 1.570796, 1.822182],accel_mss,speed_ms,0,blend_radius_m)
  movel([0.251326, -1.402353, -2.537305, -0.772731, 1.570796, 1.822122],accel_mss,speed_ms,0,blend_radius_m)
  movel([0.251281, -1.402080, -2.537508, -0.772801, 1.570796, 1.822077],accel_mss,speed_ms,0,blend_radius_m)
  movel([0.251247, -1.401798, -2.537717, -0.772874, 1.570796, 1.822043],accel_mss,speed_ms,0,blend_radius_m)
  movel([0.251229, -1.401548, -2.537902, -0.772939, 1.570796, 1.822025],accel_mss,speed_ms,0,blend_radius_m)
  movel([0.251228, -1.401291, -2.538093, -0.773005, 1.570796, 1.822025],accel_mss,speed_ms,0,blend_radius_m)
  movel([0.251243, -1.401030, -2.538286, -0.773073, 1.570796, 1.822039],accel_mss,speed_ms,0,blend_radius_m)
  movel([0.251276, -1.400741, -2.538500, -0.773148, 1.570796, 1.822072],accel_mss,speed_ms,0,blend_radius_m)
  movel([0.251323, -1.400450, -2.538715, -0.773223, 1.570796, 1.822119],accel_mss,speed_ms,0,blend_radius_m)
  movel([0.251384, -1.400157, -2.538932, -0.773300, 1.570796, 1.822180],accel_mss,speed_ms,0,blend_radius_m)
  movel([0.251482, -1.399772, -2.539217, -0.773400, 1.570796, 1.822278],accel_mss,speed_ms,0,blend_radius_m)
  movel([0.251585, -1.399386, -2.539502, -0.773501, 1.570796, 1.822381],accel_mss,speed_ms,0,blend_radius_m)
  movel([0.251699, -1.399000, -2.539786, -0.773602, 1.570796, 1.822495],accel_mss,speed_ms,0,blend_radius_m)
  movel([0.251879, -1.398424, -2.540211, -0.773754, 1.570796, 1.822675],accel_mss,speed_ms,0,blend_radius_m)
  movel([0.252046, -1.397929, -2.540576, -0.773884, 1.570796, 1.822842],accel_mss,speed_ms,0,blend_radius_m)
  movel([0.252194, -1.397502, -2.540890, -0.773997, 1.570796, 1.822991],accel_mss,speed_ms,0,blend_radius_m)
  movel([0.252213, -1.397468, -2.540915, -0.774006, 1.570796, 1.823009],accel_mss,speed_ms,0,blend_radius_m)
  movel([0.252239, -1.397440, -2.540936, -0.774013, 1.570796, 1.823035],accel_mss,speed_ms,0,blend_radius_m)
  movel([0.252263, -1.397426, -2.540946, -0.774017, 1.570796, 1.823059],accel_mss,speed_ms,0,blend_radius_m)
  movel([0.252288, -1.397417, -2.540953, -0.774020, 1.570796, 1.823084],accel_mss,speed_ms,0,blend_radius_m)
  movel([0.252311, -1.397415, -2.540954, -0.774020, 1.570796, 1.823107],accel_mss,speed_ms,0,blend_radius_m)
  movel([0.256557, -1.397998, -2.540525, -0.773866, 1.570796, 1.827354],accel_mss,speed_ms,0,blend_radius_m)
  movel([0.261236, -1.398677, -2.540025, -0.773687, 1.570796, 1.832032],accel_mss,speed_ms,0,blend_radius_m)
  movel([0.266759, -1.399523, -2.539400, -0.773465, 1.570796, 1.837555],accel_mss,speed_ms,0,blend_radius_m)
  movel([0.272287, -1.400416, -2.538741, -0.773232, 1.570796, 1.843084],accel_mss,speed_ms,0,blend_radius_m)
  movel([0.277015, -1.401209, -2.538154, -0.773026, 1.570796, 1.847812],accel_mss,speed_ms,0,blend_radius_m)
  movel([0.281147, -1.401924, -2.537623, -0.772841, 1.570796, 1.851943],accel_mss,speed_ms,0,blend_radius_m)
  movel([0.281794, -1.402042, -2.537536, -0.772811, 1.570796, 1.852590],accel_mss,speed_ms,0,blend_radius_m)
  movel([0.281967, -1.402090, -2.537500, -0.772799, 1.570796, 1.852763],accel_mss,speed_ms,0,blend_radius_m)
  speed_ms = 0.003
  movel([0.281967, -1.389907, -2.531555, -0.790927, 1.570796, 1.852763],accel_mss,speed_ms,0,blend_radius_m)
  speed_ms = 0.01
  movel([0.281967, -1.366505, -2.519283, -0.826601, 1.570796, 1.852763],accel_mss,speed_ms,0,blend_radius_m)
  movel([0.275139, -1.351369, -2.529790, -0.831230, 1.570796, 1.845936],accel_mss,speed_ms,0,blend_radius_m)
  movel([0.275139, -1.375017, -2.542249, -0.795123, 1.570796, 1.845936],accel_mss,speed_ms,0,blend_radius_m)
  speed_ms = 0.003
  movel([0.275139, -1.384229, -2.546791, -0.781369, 1.570796, 1.845936],accel_mss,speed_ms,0,blend_radius_m)
  speed_ms = 0.007
  movel([0.275100, -1.384253, -2.546774, -0.781362, 1.570796, 1.845897],accel_mss,speed_ms,0,blend_radius_m)
  movel([0.275061, -1.384262, -2.546767, -0.781359, 1.570796, 1.845858],accel_mss,speed_ms,0,blend_radius_m)
  movel([0.274454, -1.384304, -2.546737, -0.781348, 1.570796, 1.845251],accel_mss,speed_ms,0,blend_radius_m)
  movel([0.273756, -1.384340, -2.546712, -0.781338, 1.570796, 1.844552],accel_mss,speed_ms,0,blend_radius_m)
  movel([0.272946, -1.384368, -2.546691, -0.781330, 1.570796, 1.843742],accel_mss,speed_ms,0,blend_radius_m)
  movel([0.270848, -1.384429, -2.546647, -0.781312, 1.570796, 1.841644],accel_mss,speed_ms,0,blend_radius_m)
  movel([0.270977, -1.384094, -2.546888, -0.781407, 1.570796, 1.841773],accel_mss,speed_ms,0,blend_radius_m)
  movel([0.271720, -1.382154, -2.548277, -0.781958, 1.570796, 1.842517],accel_mss,speed_ms,0,blend_radius_m)
  movel([0.278710, -1.364143, -2.560921, -0.787325, 1.570796, 1.849506],accel_mss,speed_ms,0,blend_radius_m)
  movel([0.285537, -1.346758, -2.572700, -0.792931, 1.570796, 1.856333],accel_mss,speed_ms,0,blend_radius_m)
  movel([0.287626, -1.341486, -2.576190, -0.794713, 1.570796, 1.858423],accel_mss,speed_ms,0,blend_radius_m)
  movel([0.289808, -1.335986, -2.579792, -0.796612, 1.570796, 1.860604],accel_mss,speed_ms,0,blend_radius_m)
  movel([0.289826, -1.335965, -2.579805, -0.796619, 1.570796, 1.860622],accel_mss,speed_ms,0,blend_radius_m)
  movel([0.289853, -1.335945, -2.579818, -0.796626, 1.570796, 1.860650],accel_mss,speed_ms,0,blend_radius_m)
  movel([0.289881, -1.335933, -2.579826, -0.796630, 1.570796, 1.860678],accel_mss,speed_ms,0,blend_radius_m)
  movel([0.289919, -1.335919, -2.579835, -0.796635, 1.570796, 1.860715],accel_mss,speed_ms,0,blend_radius_m)
  movel([0.289955, -1.335912, -2.579840, -0.796638, 1.570796, 1.860751],accel_mss,speed_ms,0,blend_radius_m)
  movel([0.290037, -1.335908, -2.579842, -0.796639, 1.570796, 1.860833],accel_mss,speed_ms,0,blend_radius_m)
  movel([0.294408, -1.335800, -2.579912, -0.796677, 1.570796, 1.865205],accel_mss,speed_ms,0,blend_radius_m)
  movel([0.294728, -1.335799, -2.579913, -0.796677, 1.570796, 1.865524],accel_mss,speed_ms,0,blend_radius_m)
  movel([0.295043, -1.335812, -2.579904, -0.796672, 1.570796, 1.865839],accel_mss,speed_ms,0,blend_radius_m)
  movel([0.295202, -1.335829, -2.579894, -0.796667, 1.570796, 1.865998],accel_mss,speed_ms,0,blend_radius_m)
  movel([0.295351, -1.335863, -2.579871, -0.796655, 1.570796, 1.866147],accel_mss,speed_ms,0,blend_radius_m)
  movel([0.295384, -1.335880, -2.579861, -0.796649, 1.570796, 1.866180],accel_mss,speed_ms,0,blend_radius_m)
